{region "05 - Child 1 completes despite the held helper error"}
FSteps[5].Children[1].State := E_State.Completed;
FSteps[5].Children[1].Ready := FALSE;
FSteps[5].Children[1].Complete := TRUE;
FSteps[5].Children[1].Result := E_Result.Passed;
FSteps[5].Children[2].State := E_State.Idle;
FSteps[5].Children[2].Ready := FALSE;
FSteps[5].ExpectedSlot := 1;
FSteps[5].ExpectedReservations[1] := 1;
FSteps[5].MaxActiveChildCount := 1;
FSteps[5].ExpectedResult := E_Result.Error;
FSteps[5].ExpectedDiagnosticCount := 1;
{endregion}

{region "06 - Release the completed child only"}
FSteps[6].Children[1].State := E_State.Completed;
FSteps[6].Children[1].Ready := FALSE;
FSteps[6].Children[1].Complete := TRUE;
FSteps[6].Children[1].Result := E_Result.Passed;
FSteps[6].Children[2].State := E_State.Idle;
FSteps[6].Children[2].Ready := FALSE;
FSteps[6].ExpectedSlot := 1;
FSteps[6].ExpectedReleasedEntries[1] := 1;
FSteps[6].MaxActiveChildCount := 0;
FSteps[6].ExpectedResult := E_Result.Error;
FSteps[6].ExpectedDiagnosticCount := 1;
{endregion}

{region "07 - Readiness recovery does not clear the held error"}
FSteps[7].Children[1].State := E_State.Completed;
FSteps[7].Children[1].Ready := FALSE;
FSteps[7].Children[1].Complete := TRUE;
FSteps[7].Children[1].Result := E_Result.Passed;
FSteps[7].ExpectedSlot := 1;
FSteps[7].MaxActiveChildCount := 0;
FSteps[7].ExpectedResult := E_Result.Error;
FSteps[7].ExpectedDiagnosticCount := 1;
{endregion}

{region "08 - Recovered readiness cannot restart execution"}
FSteps[8].Children[1].State := E_State.Completed;
FSteps[8].Children[1].Ready := FALSE;
FSteps[8].Children[1].Complete := TRUE;
FSteps[8].Children[1].Result := E_Result.Passed;
FSteps[8].ExpectedSlot := 1;
FSteps[8].MaxActiveChildCount := 0;
FSteps[8].ExpectedResult := E_Result.Error;
FSteps[8].ExpectedDiagnosticCount := 1;
{endregion}
END_METHOD

END_FUNCTION_BLOCK

// ---- SelfTests/TestCases/TestSuite_ParallelOrchestration/Test_ParallelFailedResultContinues.TcPOU
{region 'Documentation'}
(*!
<summary>Keeps parallel siblings progressing after a child completes with Failed instead of treating it as a helper Error.</summary>
<description>
Child 1 finishes with Failed while child 2 starts. Child 3 must still start while child 2
runs. The helper reports neutral Result and completes only after all children;
child-result aggregation belongs to the owner.
</description>
*)
{endregion}
FUNCTION_BLOCK Test_ParallelFailedResultContinues EXTENDS OrchestrationTestBase

SUPER^();

{region 'Documentation'}
(*!
<summary>Defines reachable child responses and independent per-cycle expectations.</summary>
*)
{endregion}
METHOD PROTECTED ConfigureScenario
FChildSlots[1] := 1;
FChildSlots[2] := 1;
FChildSlots[3] := 1;
FStepCount := 7;

{region "01 - Observe initial readiness"}
FSteps[1].Task := E_OrchestratorTask.Idle;
FSteps[1].ExpectedReady := TRUE;
{endregion}

{region "02 - Start child 1"}
FSteps[2].Children[1].State := E_State.Running;
FSteps[2].Children[1].Ready := FALSE;
FSteps[2].ExpectedStartChild := 1;
FSteps[2].ExpectedSlot := 1;
FSteps[2].ExpectedReservations[1] := 1;
FSteps[2].MaxActiveChildCount := 1;
{endregion}

{region "03 - Start child 2 while child 1 finishes with Failed"}
FSteps[3].Children[1].State := E_State.Completed;
FSteps[3].Children[1].Ready := FALSE;
FSteps[3].Children[1].Complete := TRUE;
FSteps[3].Children[1].Result := E_Result.Failed;
FSteps[3].Children[2].State := E_State.Running;
FSteps[3].Children[2].Ready := FALSE;
FSteps[3].ExpectedStartChild := 2;
FSteps[3].ExpectedSlot := 1;
FSteps[3].ExpectedReservations[1] := 1;
FSteps[3].ExpectedReservations[2] := 1;
FSteps[3].MaxActiveChildCount := 2;
{endregion}

{region "04 - Release Failed child 1 and start child 3"}
FSteps[4].Children[1].State := E_State.Completed;
FSteps[4].Children[1].Ready := FALSE;
FSteps[4].Children[1].Complete := TRUE;
FSteps[4].Children[1].Result := E_Result.Failed;
FSteps[4].Children[2].State := E_State.Running;
FSteps[4].Children[2].Ready := FALSE;
FSteps[4].Children[3].State := E_State.Running;
FSteps[4].Children[3].Ready := FALSE;
FSteps[4].ExpectedStartChild := 3;
FSteps[4].ExpectedSlot := 1;
FSteps[4].ExpectedReservations[2] := 1;
FSteps[4].ExpectedReservations[3] := 1;
FSteps[4].ExpectedReleasedEntries[1] := 1;
FSteps[4].MaxActiveChildCount := 2;
{endregion}

{region "05 - Remaining children complete without helper Error"}
FSteps[5].Children[1].State := E_State.Completed;
FSteps[5].Children[1].Ready := FALSE;
FSteps[5].Children[1].Complete := TRUE;
FSteps[5].Children[1].Result := E_Result.Failed;
FSteps[5].Children[2].State := E_State.Completed;
FSteps[5].Children[2].Ready := FALSE;
FSteps[5].Children[2].Complete := TRUE;
FSteps[5].Children[2].Result := E_Result.Passed;
FSteps[5].Children[3].State := E_State.Completed;
FSteps[5].Children[3].Ready := FALSE;
FSteps[5].Children[3].Complete := TRUE;
FSteps[5].Children[3].Result := E_Result.Passed;
FSteps[5].ExpectedSlot := 1;
FSteps[5].ExpectedReservations[2] := 1;
FSteps[5].ExpectedReservations[3] := 1;
FSteps[5].MaxActiveChildCount := 2;
{endregion}

{region "06 - Release both siblings and finish the whole group"}
FSteps[6].Children[1].State := E_State.Completed;
FSteps[6].Children[1].Ready := FALSE;
FSteps[6].Children[1].Complete := TRUE;
FSteps[6].Children[1].Result := E_Result.Failed;
FSteps[6].Children[2].State := E_State.Completed;
FSteps[6].Children[2].Ready := FALSE;
FSteps[6].Children[2].Complete := TRUE;
FSteps[6].Children[2].Result := E_Result.Passed;
FSteps[6].Children[3].State := E_State.Completed;
FSteps[6].Children[3].Ready := FALSE;
FSteps[6].Children[3].Complete := TRUE;
FSteps[6].Children[3].Result := E_Result.Passed;
FSteps[6].ExpectedFinished := TRUE;
FSteps[6].ExpectedReleasedEntries[2] := 1;
FSteps[6].ExpectedReleasedEntries[3] := 1;
FSteps[6].MaxActiveChildCount := 0;
{endregion}

{region "07 - Keep completion stable with neutral helper Result"}
FSteps[7].Children[1].State := E_State.Completed;
FSteps[7].Children[1].Ready := FALSE;
FSteps[7].Children[1].Complete := TRUE;
FSteps[7].Children[1].Result := E_Result.Failed;
FSteps[7].Children[2].State := E_State.Completed;
FSteps[7].Children[2].Ready := FALSE;
FSteps[7].Children[2].Complete := TRUE;
FSteps[7].Children[2].Result := E_Result.Passed;
FSteps[7].Children[3].State := E_State.Completed;
FSteps[7].Children[3].Ready := FALSE;
FSteps[7].Children[3].Complete := TRUE;
FSteps[7].Children[3].Result := E_Result.Passed;
FSteps[7].ExpectedFinished := TRUE;
FSteps[7].MaxActiveChildCount := 0;
{endregion}
END_METHOD

END_FUNCTION_BLOCK

// ---- SelfTests/TestCases/TestSuite_ParallelOrchestration/Test_ParallelChildError.TcPOU
{region 'Documentation'}
(*!
<summary>Stops new parallel Starts on child Error and observes owner-selected Abort of the remaining active sibling.</summary>
<description>
Child 1 enters its error-abort path while child 2 starts. The helper must retain Error and
not start child 3. The owner then supplies Abort explicitly; already-aborting child 1 and
never-started child 3 receive no redundant Abort.
</description>
*)
{endregion}
FUNCTION_BLOCK Test_ParallelChildError EXTENDS OrchestrationTestBase

SUPER^();

{region 'Documentation'}
(*!
<summary>Defines reachable child responses and independent per-cycle expectations.</summary>
*)
{endregion}
METHOD PROTECTED ConfigureScenario
FChildSlots[1] := 1;
FChildSlots[2] := 1;
FChildSlots[3] := 1;
FStepCount := 8;

{region "01 - Observe initial readiness"}
FSteps[1].Task := E_OrchestratorTask.Idle;
FSteps[1].ExpectedReady := TRUE;
{endregion}

{region "02 - Start child 1 normally"}
FSteps[2].Children[1].State := E_State.Running;
FSteps[2].Children[1].Ready := FALSE;
FSteps[2].ExpectedStartChild := 1;
FSteps[2].ExpectedSlot := 1;
FSteps[2].ExpectedReservations[1] := 1;
FSteps[2].MaxActiveChildCount := 1;
{endregion}

{region "03 - Start child 2 while child 1 enters its error path"}
FSteps[3].Children[1].State := E_State.AbortingFromError;
FSteps[3].Children[1].Ready := FALSE;
FSteps[3].Children[1].Result := E_Result.Error;
FSteps[3].Children[2].State := E_State.Running;
FSteps[3].Children[2].Ready := FALSE;
FSteps[3].ExpectedStartChild := 2;
FSteps[3].ExpectedSlot := 1;
FSteps[3].ExpectedReservations[1] := 1;
FSteps[3].ExpectedReservations[2] := 1;
FSteps[3].MaxActiveChildCount := 2;
{endregion}

{region "04 - Observe child Error and suppress child 3 Start"}
FSteps[4].Children[1].State := E_State.AbortingFromError;
FSteps[4].Children[1].Ready := FALSE;
FSteps[4].Children[1].Result := E_Result.Error;
FSteps[4].Children[2].State := E_State.Running;
FSteps[4].Children[2].Ready := FALSE;
FSteps[4].ExpectedSlot := 1;
FSteps[4].ExpectedReservations[1] := 1;
FSteps[4].ExpectedReservations[2] := 1;
FSteps[4].MaxActiveChildCount := 2;
FSteps[4].ExpectedResult := E_Result.Error;
FSteps[4].ExpectedDiagnosticCount := 1;
{endregion}

{region "05 - Owner selects Abort for remaining active work"}
FSteps[5].Task := E_OrchestratorTask.Abort;
FSteps[5].Children[1].State := E_State.AbortingFromError;
FSteps[5].Children[1].Ready := FALSE;
FSteps[5].Children[1].Result := E_Result.Error;
FSteps[5].Children[2].State := E_State.Aborting;
FSteps[5].Children[2].Ready := FALSE;
FSteps[5].Children[2].Result := E_Result.Abort;
FSteps[5].ExpectedReservations[1] := 1;
FSteps[5].ExpectedReservations[2] := 1;
FSteps[5].ExpectedAbortRequests[2] := 1;
FSteps[5].ExpectedResult := E_Result.Error;
FSteps[5].ExpectedDiagnosticCount := 1;
{endregion}

{region "06 - Both active children reach terminal states"}
FSteps[6].Task := E_OrchestratorTask.Abort;
FSteps[6].Children[1].State := E_State.Completed;
FSteps[6].Children[1].Ready := FALSE;
FSteps[6].Children[1].Complete := TRUE;
FSteps[6].Children[1].Result := E_Result.Error;
FSteps[6].Children[2].State := E_State.Completed;
FSteps[6].Children[2].Ready := FALSE;
FSteps[6].Children[2].Complete := TRUE;
FSteps[6].Children[2].Result := E_Result.Abort;
FSteps[6].ExpectedReservations[1] := 1;
FSteps[6].ExpectedReservations[2] := 1;
FSteps[6].ExpectedResult := E_Result.Error;
FSteps[6].ExpectedDiagnosticCount := 1;
{endregion}

{region "07 - Release terminal reservations and finish Abort"}
FSteps[7].Task := E_OrchestratorTask.Abort;
FSteps[7].Children[1].State := E_State.Completed;
FSteps[7].Children[1].Ready := FALSE;
FSteps[7].Children[1].Complete := TRUE;
FSteps[7].Children[1].Result := E_Result.Error;
FSteps[7].Children[2].State := E_State.Completed;
FSteps[7].Children[2].Ready := FALSE;
FSteps[7].Children[2].Complete := TRUE;
FSteps[7].Children[2].Result := E_Result.Abort;
FSteps[7].ExpectedAbortFinished := TRUE;
FSteps[7].ExpectedReleasedEntries[1] := 1;
FSteps[7].ExpectedReleasedEntries[2] := 1;
FSteps[7].ExpectedResult := E_Result.Error;
FSteps[7].ExpectedDiagnosticCount := 1;
{endregion}

{region "08 - Repeated Abort neither redispatches nor republishes"}
FSteps[8].Task := E_OrchestratorTask.Abort;
FSteps[8].Children[1].State := E_State.Completed;
FSteps[8].Children[1].Ready := FALSE;
FSteps[8].Children[1].Complete := TRUE;
FSteps[8].Children[1].Result := E_Result.Error;
FSteps[8].Children[2].State := E_State.Completed;
FSteps[8].Children[2].Ready := FALSE;
FSteps[8].Children[2].Complete := TRUE;
FSteps[8].Children[2].Result := E_Result.Abort;
FSteps[8].ExpectedAbortFinished := TRUE;
FSteps[8].ExpectedResult := E_Result.Error;
FSteps[8].ExpectedDiagnosticCount := 1;
{endregion}
END_METHOD

END_FUNCTION_BLOCK

// ---- SelfTests/TestCases/TestSuite_ParallelOrchestration/Test_ParallelAbortMixedProgress.TcPOU
{region 'Documentation'}
(*!
<summary>Aborts only active parallel work while leaving completed and never-started ready children untouched.</summary>
<description>
Child 2 completes on its Start call while child 1 runs. The owner selects Abort before
child 3 starts. Start confirmation, terminal release and active-child Abort happen in the
same helper call; completion waits for child 1.
</description>
*)
{endregion}
FUNCTION_BLOCK Test_ParallelAbortMixedProgress EXTENDS OrchestrationTestBase

SUPER^();

{region 'Documentation'}
(*!
<summary>Defines reachable child responses and independent per-cycle expectations.</summary>
*)
{endregion}
METHOD PROTECTED ConfigureScenario
FChildSlots[1] := 1;
FChildSlots[2] := 1;
FChildSlots[3] := 1;
FStepCount := 7;

{region "01 - Observe initial readiness"}
FSteps[1].Task := E_OrchestratorTask.Idle;
FSteps[1].ExpectedReady := TRUE;
{endregion}

{region "02 - Start child 1"}
FSteps[2].Children[1].State := E_State.Running;
FSteps[2].Children[1].Ready := FALSE;
FSteps[2].ExpectedStartChild := 1;
FSteps[2].ExpectedSlot := 1;
FSteps[2].ExpectedReservations[1] := 1;
FSteps[2].MaxActiveChildCount := 1;
{endregion}

{region "03 - Start immediately completing child 2"}
FSteps[3].Children[1].State := E_State.Running;
FSteps[3].Children[1].Ready := FALSE;
FSteps[3].Children[2].State := E_State.Completed;
FSteps[3].Children[2].Ready := FALSE;
FSteps[3].Children[2].Complete := TRUE;
FSteps[3].Children[2].Result := E_Result.Passed;
FSteps[3].ExpectedStartChild := 2;
FSteps[3].ExpectedSlot := 1;
FSteps[3].ExpectedReservations[1] := 1;
FSteps[3].ExpectedReservations[2] := 1;
FSteps[3].MaxActiveChildCount := 2;
{endregion}

{region "04 - Owner selects Abort while child 3 remains unstarted"}
FSteps[4].Task := E_OrchestratorTask.Abort;
FSteps[4].Children[1].State := E_State.Aborting;
FSteps[4].Children[1].Ready := FALSE;
FSteps[4].Children[1].Result := E_Result.Abort;
FSteps[4].Children[2].State := E_State.Completed;
FSteps[4].Children[2].Ready := FALSE;
FSteps[4].Children[2].Complete := TRUE;
FSteps[4].Children[2].Result := E_Result.Passed;
FSteps[4].ExpectedReservations[1] := 1;
FSteps[4].ExpectedReleasedEntries[2] := 1;
FSteps[4].ExpectedAbortRequests[1] := 1;
{endregion}

{region "05 - Wait for the active child's controlled completion"}
FSteps[5].Task := E_OrchestratorTask.Abort;
FSteps[5].Children[1].State := E_State.Completed;
FSteps[5].Children[1].Ready := FALSE;
FSteps[5].Children[1].Complete := TRUE;
FSteps[5].Children[1].Result := E_Result.Abort;
FSteps[5].Children[2].State := E_State.Completed;
FSteps[5].Children[2].Ready := FALSE;
FSteps[5].Children[2].Complete := TRUE;
FSteps[5].Children[2].Result := E_Result.Passed;
FSteps[5].ExpectedReservations[1] := 1;
{endregion}

{region "06 - Release child 1 and finish Abort"}
FSteps[6].Task := E_OrchestratorTask.Abort;
FSteps[6].Children[1].State := E_State.Completed;
FSteps[6].Children[1].Ready := FALSE;
FSteps[6].Children[1].Complete := TRUE;
FSteps[6].Children[1].Result := E_Result.Abort;
FSteps[6].Children[2].State := E_State.Completed;
FSteps[6].Children[2].Ready := FALSE;
FSteps[6].Children[2].Complete := TRUE;
FSteps[6].Children[2].Result := E_Result.Passed;
FSteps[6].ExpectedAbortFinished := TRUE;
FSteps[6].ExpectedReleasedEntries[1] := 1;
{endregion}

{region "07 - No repeated Abort or new Start after completion"}
FSteps[7].Task := E_OrchestratorTask.Abort;
FSteps[7].Children[1].State := E_State.Completed;
FSteps[7].Children[1].Ready := FALSE;
FSteps[7].Children[1].Complete := TRUE;
FSteps[7].Children[1].Result := E_Result.Abort;
FSteps[7].Children[2].State := E_State.Completed;
FSteps[7].Children[2].Ready := FALSE;
FSteps[7].Children[2].Complete := TRUE;
FSteps[7].Children[2].Result := E_Result.Passed;
FSteps[7].ExpectedAbortFinished := TRUE;
{endregion}
END_METHOD

END_FUNCTION_BLOCK

// ---- SelfTests/TestCases/TestSuite_ParallelOrchestration/Test_ParallelResetOverlappingExecution.TcPOU
{region 'Documentation'}
(*!
<summary>Resets overlapping parallel children and an already completed child without issuing further Starts.</summary>
<description>
Two children are running when the third completes immediately. Owner-selected Reset
replaces each execution reservation through the child's Reset reservation method.
Independent reset completion retains unfinished reservations and returns to ready Idle
only after all children finish.
</description>
*)
{endregion}
FUNCTION_BLOCK Test_ParallelResetOverlappingExecution EXTENDS OrchestrationTestBase

SUPER^();

{region 'Documentation'}
(*!
<summary>Defines reachable child responses and independent per-cycle expectations.</summary>
*)
{endregion}
METHOD PROTECTED ConfigureScenario
FChildSlots[1] := 1;
FChildSlots[2] := 1;
FChildSlots[3] := 1;
FStepCount := 12;

{region "01 - Observe initial readiness"}
FSteps[1].Task := E_OrchestratorTask.Idle;
FSteps[1].ExpectedReady := TRUE;
{endregion}

{region "02 - Start child 1"}
FSteps[2].Children[1].State := E_State.Running;
FSteps[2].Children[1].Ready := FALSE;
FSteps[2].ExpectedStartChild := 1;
FSteps[2].ExpectedSlot := 1;
FSteps[2].ExpectedReservations[1] := 1;
FSteps[2].MaxActiveChildCount := 1;
{endregion}

{region "03 - Start child 2 concurrently"}
FSteps[3].Children[1].State := E_State.Running;
FSteps[3].Children[1].Ready := FALSE;
FSteps[3].Children[2].State := E_State.Running;
FSteps[3].Children[2].Ready := FALSE;
FSteps[3].ExpectedStartChild := 2;
FSteps[3].ExpectedSlot := 1;
FSteps[3].ExpectedReservations[1] := 1;
FSteps[3].ExpectedReservations[2] := 1;
FSteps[3].MaxActiveChildCount := 2;
{endregion}

{region "04 - Start child 3 which completes immediately"}
FSteps[4].Children[1].State := E_State.Running;
FSteps[4].Children[1].Ready := FALSE;
FSteps[4].Children[2].State := E_State.Running;
FSteps[4].Children[2].Ready := FALSE;
FSteps[4].Children[3].State := E_State.Completed;
FSteps[4].Children[3].Ready := FALSE;
FSteps[4].Children[3].Complete := TRUE;
FSteps[4].Children[3].Result := E_Result.Passed;
FSteps[4].ExpectedStartChild := 3;
FSteps[4].ExpectedSlot := 1;
FSteps[4].ExpectedReservations[1] := 1;
FSteps[4].ExpectedReservations[2] := 1;
FSteps[4].ExpectedReservations[3] := 1;
FSteps[4].MaxActiveChildCount := 3;
{endregion}

{region "05 - Owner selects Reset and resets active child 1"}
FSteps[5].Task := E_OrchestratorTask.Reset;
FSteps[5].Children[1].State := E_State.Reset;
FSteps[5].Children[1].Ready := FALSE;
FSteps[5].Children[2].State := E_State.Running;
FSteps[5].Children[2].Ready := FALSE;
FSteps[5].Children[3].State := E_State.Completed;
FSteps[5].Children[3].Ready := FALSE;
FSteps[5].Children[3].Complete := TRUE;
FSteps[5].Children[3].Result := E_Result.Passed;
FSteps[5].ExpectedResetChild := 1;
FSteps[5].ExpectedReservations[1] := 1;
FSteps[5].ExpectedReservations[2] := 1;
FSteps[5].ExpectedReservations[3] := 1;
{endregion}

{region "06 - Reset child 2 while child 1 is still resetting"}
FSteps[6].Task := E_OrchestratorTask.Reset;
FSteps[6].Children[1].State := E_State.Reset;
FSteps[6].Children[1].Ready := FALSE;
FSteps[6].Children[2].State := E_State.Reset;
FSteps[6].Children[2].Ready := FALSE;
FSteps[6].Children[3].State := E_State.Completed;
FSteps[6].Children[3].Ready := FALSE;
FSteps[6].Children[3].Complete := TRUE;
FSteps[6].Children[3].Result := E_Result.Passed;
FSteps[6].ExpectedResetChild := 2;
FSteps[6].ExpectedReservations[1] := 1;
FSteps[6].ExpectedReservations[2] := 1;
FSteps[6].ExpectedReservations[3] := 1;
{endregion}

{region "07 - Reset completed child 3 while child 1 reaches Idle"}
FSteps[7].Task := E_OrchestratorTask.Reset;
FSteps[7].Children[2].State := E_State.Reset;
FSteps[7].Children[2].Ready := FALSE;
FSteps[7].Children[3].State := E_State.Reset;
FSteps[7].Children[3].Ready := FALSE;
FSteps[7].ExpectedResetChild := 3;
FSteps[7].ExpectedReservations[1] := 1;
FSteps[7].ExpectedReservations[2] := 1;
FSteps[7].ExpectedReservations[3] := 1;
{endregion}

{region "08 - Release child 1 while child 2 reaches Idle"}
FSteps[8].Task := E_OrchestratorTask.Reset;
FSteps[8].Children[3].State := E_State.Reset;
FSteps[8].Children[3].Ready := FALSE;
FSteps[8].ExpectedReservations[2] := 1;
FSteps[8].ExpectedReservations[3] := 1;
FSteps[8].ExpectedReleasedEntries[1] := 1;
{endregion}

{region "09 - Release child 2 while child 3 reaches Idle"}
FSteps[9].Task := E_OrchestratorTask.Reset;
FSteps[9].ExpectedReservations[3] := 1;
FSteps[9].ExpectedReleasedEntries[2] := 1;
{endregion}

{region "10 - Release final reservation and report Reset finished"}
FSteps[10].Task := E_OrchestratorTask.Reset;
FSteps[10].ExpectedResetFinished := TRUE;
FSteps[10].ExpectedReleasedEntries[3] := 1;
{endregion}

{region "11 - Repeated Reset retains completion without redispatch"}
FSteps[11].Task := E_OrchestratorTask.Reset;
FSteps[11].ExpectedResetFinished := TRUE;
{endregion}

{region "12 - Owner selects Idle and observes restored readiness"}
FSteps[12].Task := E_OrchestratorTask.Idle;
FSteps[12].ExpectedReady := TRUE;
{endregion}
END_METHOD

END_FUNCTION_BLOCK

// ---- SelfTests/TestSuites/TestSuite_ParallelSlotsOrchestration.TcPOU
{region 'Documentation'}
(*!
<summary>Runs focused ParallelSlots Orchestrator scenarios serially with isolated child observations and diagnostics.</summary>
*)
{endregion}
FUNCTION_BLOCK TestSuite_ParallelSlotsOrchestration EXTENDS TestSuiteBase
VAR
    FWaitForGroupCompletion : Test_SlotsWaitForGroupCompletion;
    FFinalGroupCompletion : Test_SlotsFinalGroupCompletion;
    FFirstFittingAdmission : Test_SlotsFirstFittingAdmission;
    FMissingStartReaction : Test_SlotsMissingStartReaction;
    FNextSlotReadinessLost : Test_SlotsNextSlotReadinessLost;
    FAbortAtBoundary : Test_SlotsAbortAtBoundary;
    FTestCases : ARRAY[1..TestCaseCapacity] OF I_TestCase;
END_VAR
VAR CONSTANT
    TestCaseCapacity : UINT := 6;
END_VAR

SUPER^();

{region 'Documentation'}
(*!
<summary>Initializes and registers the owned orchestration scenarios in deterministic order.</summary>
*)
{endregion}
METHOD PROTECTED Configure
VAR_IN_OUT
    // SA0167: Borrowed builder; VAR_IN_OUT creates no temporary instance.
    {attribute 'analysis' := '-167'}
    Builder : TestSuiteConfigurationBuilder; //! Borrowed owner configuration builder used only during this Configure call; register this owner's concrete children.
END_VAR
VAR
    TestConfig : ST_TestCaseConfig;
END_VAR
Builder.Initialize(Mode := E_OrchestrationMode.Serial,
    TestCases := FTestCases);

FWaitForGroupCompletion.Initialize(Parent := THIS^,
    TestName := 'WaitForGroupCompletion',
    Config := TestConfig);
Builder.Register(TestCase := FWaitForGroupCompletion);

FFinalGroupCompletion.Initialize(Parent := THIS^,
    TestName := 'FinalGroupCompletion',
    Config := TestConfig);
Builder.Register(TestCase := FFinalGroupCompletion);

FFirstFittingAdmission.Initialize(Parent := THIS^,
    TestName := 'FirstFittingAdmission',
    Config := TestConfig);
Builder.Register(TestCase := FFirstFittingAdmission);

FMissingStartReaction.Initialize(Parent := THIS^,
    TestName := 'MissingStartReaction',
    Config := TestConfig);
Builder.Register(TestCase := FMissingStartReaction);

FNextSlotReadinessLost.Initialize(Parent := THIS^,
    TestName := 'NextSlotReadinessLost',
    Config := TestConfig);
Builder.Register(TestCase := FNextSlotReadinessLost);

FAbortAtBoundary.Initialize(Parent := THIS^,
    TestName := 'AbortAtBoundary',
    Config := TestConfig);
Builder.Register(TestCase := FAbortAtBoundary);
END_METHOD

{region 'Documentation'}
(*!
<summary>Returns the registered Test Case from the same array used during configuration.</summary>
*)
{endregion}
METHOD PUBLIC GetTestCase : I_TestCase //! Typed child interface at the original array index; zero when no entry is available.
VAR_INPUT
    Index : DINT; //! Original occupied child-array index, rather than an ordinal position.
END_VAR
GetTestCase := 0;
IF (ChildCount = 0) OR (Index < ChildArrayLowerBound)
    OR (DINT_TO_LINT(Index) >= DINT_TO_LINT(ChildArrayLowerBound) + UINT_TO_LINT(ChildCount)) THEN
    RETURN;
END_IF;

GetTestCase := FTestCases[Index];
END_METHOD

{region 'Documentation'}
(*!
<summary>Calls each owned Test Case once per initialized Suite cycle, including completion.</summary>
*)
{endregion}
METHOD PROTECTED ProcessTestCases
FWaitForGroupCompletion();
FFinalGroupCompletion();
FFirstFittingAdmission();
FMissingStartReaction();
FNextSlotReadinessLost();
FAbortAtBoundary();
END_METHOD

END_FUNCTION_BLOCK

// ---- SelfTests/TestCases/TestSuite_ParallelSlotsOrchestration/Test_SlotsWaitForGroupCompletion.TcPOU
{region 'Documentation'}
(*!
<summary>Keeps the next slot blocked until both unequal-duration children in the current slot complete.</summary>
<description>
Children 1 and 2 share slot 1. Child 2 finishes first while child 1 remains active.
Child 3 stays idle in slot 2 until both earlier children complete and their reservations
are released. Each row observes the helper before applying the next child responses.
</description>
*)
{endregion}
FUNCTION_BLOCK Test_SlotsWaitForGroupCompletion EXTENDS OrchestrationTestBase

SUPER^();

{region 'Documentation'}
(*!
<summary>Defines slot-group stimuli and per-cycle dispatch, completion and reservation expectations.</summary>
*)
{endregion}
METHOD PROTECTED ConfigureScenario
FChildSlots[1] := 1;
FChildSlots[2] := 1;
FChildSlots[3] := 2;
FStepCount := 11;

{region "01 - Observe initial readiness"}
FSteps[1].Task := E_OrchestratorTask.Idle;
FSteps[1].ExpectedReady := TRUE;
FSteps[1].MaxActiveChildCount := 0;
{endregion}

{region "02 - Start long-running child 1 in slot 1"}
FSteps[2].Children[1].State := E_State.Running;
FSteps[2].Children[1].Ready := FALSE;
FSteps[2].ExpectedStartChild := 1;
FSteps[2].ExpectedSlot := 1;
FSteps[2].ExpectedReservations[1] := 1;
FSteps[2].MaxActiveChildCount := 1;
{endregion}

{region "03 - Start child 2 alongside child 1"}
FSteps[3].Children[1].State := E_State.Running;
FSteps[3].Children[1].Ready := FALSE;
FSteps[3].Children[2].State := E_State.Running;
FSteps[3].Children[2].Ready := FALSE;
FSteps[3].ExpectedStartChild := 2;
FSteps[3].ExpectedSlot := 1;
FSteps[3].ExpectedReservations[1] := 1;
FSteps[3].ExpectedReservations[2] := 1;
FSteps[3].MaxActiveChildCount := 2;
{endregion}

{region "04 - Child 2 completes while child 1 remains active"}
FSteps[4].Children[1].State := E_State.Running;
FSteps[4].Children[1].Ready := FALSE;
FSteps[4].Children[2].State := E_State.Completed;
FSteps[4].Children[2].Ready := FALSE;
FSteps[4].Children[2].Complete := TRUE;
FSteps[4].Children[2].Result := E_Result.Passed;
FSteps[4].ExpectedSlot := 1;
FSteps[4].ExpectedReservations[1] := 1;
FSteps[4].ExpectedReservations[2] := 1;
FSteps[4].MaxActiveChildCount := 2;
{endregion}

{region "05 - Release child 2 without starting the next slot"}
FSteps[5].Children[1].State := E_State.Running;
FSteps[5].Children[1].Ready := FALSE;
FSteps[5].Children[2].State := E_State.Completed;
FSteps[5].Children[2].Ready := FALSE;
FSteps[5].Children[2].Complete := TRUE;
FSteps[5].Children[2].Result := E_Result.Passed;
FSteps[5].ExpectedSlot := 1;
FSteps[5].ExpectedReservations[1] := 1;
FSteps[5].ExpectedReleasedEntries[2] := 1;
FSteps[5].MaxActiveChildCount := 1;
{endregion}

{region "06 - Child 1 completes while child 3 still receives no Start"}
FSteps[6].Children[1].State := E_State.Completed;
FSteps[6].Children[1].Ready := FALSE;
FSteps[6].Children[1].Complete := TRUE;
FSteps[6].Children[1].Result := E_Result.Passed;
FSteps[6].Children[2].State := E_State.Completed;
FSteps[6].Children[2].Ready := FALSE;
FSteps[6].Children[2].Complete := TRUE;
FSteps[6].Children[2].Result := E_Result.Passed;
FSteps[6].ExpectedSlot := 1;
FSteps[6].ExpectedReservations[1] := 1;
FSteps[6].MaxActiveChildCount := 1;
{endregion}

{region "07 - Reconcile slot 1 and select slot 2 without dispatch"}
FSteps[7].Children[1].State := E_State.Completed;
FSteps[7].Children[1].Ready := FALSE;
FSteps[7].Children[1].Complete := TRUE;
FSteps[7].Children[1].Result := E_Result.Passed;
FSteps[7].Children[2].State := E_State.Completed;
FSteps[7].Children[2].Ready := FALSE;
FSteps[7].Children[2].Complete := TRUE;
FSteps[7].Children[2].Result := E_Result.Passed;
FSteps[7].ExpectedSlot := 2;
FSteps[7].ExpectedReleasedEntries[1] := 1;
FSteps[7].MaxActiveChildCount := 0;
{endregion}

{region "08 - Start child 3 only after the first group has finished"}
FSteps[8].Children[1].State := E_State.Completed;
FSteps[8].Children[1].Ready := FALSE;
FSteps[8].Children[1].Complete := TRUE;
FSteps[8].Children[1].Result := E_Result.Passed;
FSteps[8].Children[2].State := E_State.Completed;
FSteps[8].Children[2].Ready := FALSE;
FSteps[8].Children[2].Complete := TRUE;
FSteps[8].Children[2].Result := E_Result.Passed;
FSteps[8].Children[3].State := E_State.Running;
FSteps[8].Children[3].Ready := FALSE;
FSteps[8].ExpectedStartChild := 3;
FSteps[8].ExpectedSlot := 2;
FSteps[8].ExpectedReservations[3] := 1;
FSteps[8].MaxActiveChildCount := 1;
{endregion}

{region "09 - Last child completes without redispatching earlier children"}
FSteps[9].Children[1].State := E_State.Completed;
FSteps[9].Children[1].Ready := FALSE;
FSteps[9].Children[1].Complete := TRUE;
FSteps[9].Children[1].Result := E_Result.Passed;
FSteps[9].Children[2].State := E_State.Completed;
FSteps[9].Children[2].Ready := FALSE;
FSteps[9].Children[2].Complete := TRUE;
FSteps[9].Children[2].Result := E_Result.Passed;
FSteps[9].Children[3].State := E_State.Completed;
FSteps[9].Children[3].Ready := FALSE;
FSteps[9].Children[3].Complete := TRUE;
FSteps[9].Children[3].Result := E_Result.Passed;
FSteps[9].ExpectedSlot := 2;
FSteps[9].ExpectedReservations[3] := 1;
FSteps[9].MaxActiveChildCount := 1;
{endregion}

{region "10 - Release the last reservation and finish all slots"}
FSteps[10].Children[1].State := E_State.Completed;
FSteps[10].Children[1].Ready := FALSE;
FSteps[10].Children[1].Complete := TRUE;
FSteps[10].Children[1].Result := E_Result.Passed;
FSteps[10].Children[2].State := E_State.Completed;
FSteps[10].Children[2].Ready := FALSE;
FSteps[10].Children[2].Complete := TRUE;
FSteps[10].Children[2].Result := E_Result.Passed;
FSteps[10].Children[3].State := E_State.Completed;
FSteps[10].Children[3].Ready := FALSE;
FSteps[10].Children[3].Complete := TRUE;
FSteps[10].Children[3].Result := E_Result.Passed;
FSteps[10].ExpectedFinished := TRUE;
FSteps[10].ExpectedReleasedEntries[3] := 1;
FSteps[10].MaxActiveChildCount := 0;
{endregion}

{region "11 - Keep final completion stable without further Starts"}
FSteps[11].Children[1].State := E_State.Completed;
FSteps[11].Children[1].Ready := FALSE;
FSteps[11].Children[1].Complete := TRUE;
FSteps[11].Children[1].Result := E_Result.Passed;
FSteps[11].Children[2].State := E_State.Completed;
FSteps[11].Children[2].Ready := FALSE;
FSteps[11].Children[2].Complete := TRUE;
FSteps[11].Children[2].Result := E_Result.Passed;
FSteps[11].Children[3].State := E_State.Completed;
FSteps[11].Children[3].Ready := FALSE;
FSteps[11].Children[3].Complete := TRUE;
FSteps[11].Children[3].Result := E_Result.Passed;
FSteps[11].ExpectedFinished := TRUE;
FSteps[11].MaxActiveChildCount := 0;
{endregion}
END_METHOD

END_FUNCTION_BLOCK

// ---- SelfTests/TestCases/TestSuite_ParallelSlotsOrchestration/Test_SlotsFinalGroupCompletion.TcPOU
{region 'Documentation'}
(*!
<summary>Runs both final-slot children in parallel and ignores unused collection capacity when determining completion.</summary>
<description>
Child 1 completes immediately in slot 1. Children 2 and 3 then overlap in the final
slot and finish in reverse order. The collection has six array positions but only three
registered children; final-slot detection must use the occupied range.
</description>
*)
{endregion}
FUNCTION_BLOCK Test_SlotsFinalGroupCompletion EXTENDS OrchestrationTestBase

SUPER^();

{region 'Documentation'}
(*!
<summary>Defines slot-group stimuli and per-cycle dispatch, completion and reservation expectations.</summary>
*)
{endregion}
METHOD PROTECTED ConfigureScenario
FChildSlots[1] := 1;
FChildSlots[2] := 2;
FChildSlots[3] := 2;
FArrayLayout := E_OrchestrationArrayLayout.SpareCapacity;
FStepCount := 10;

{region "01 - Observe readiness with unused array capacity"}
FSteps[1].Task := E_OrchestratorTask.Idle;
FSteps[1].ExpectedReady := TRUE;
FSteps[1].MaxActiveChildCount := 0;
{endregion}

{region "02 - Start child 1 which completes immediately"}
FSteps[2].Children[1].State := E_State.Completed;
FSteps[2].Children[1].Ready := FALSE;
FSteps[2].Children[1].Complete := TRUE;
FSteps[2].Children[1].Result := E_Result.Passed;
FSteps[2].ExpectedStartChild := 1;
FSteps[2].ExpectedSlot := 1;
FSteps[2].ExpectedReservations[1] := 1;
FSteps[2].MaxActiveChildCount := 1;
{endregion}

{region "03 - Confirm immediate completion and select the final slot"}
FSteps[3].Children[1].State := E_State.Completed;
FSteps[3].Children[1].Ready := FALSE;
FSteps[3].Children[1].Complete := TRUE;
FSteps[3].Children[1].Result := E_Result.Passed;
FSteps[3].ExpectedSlot := 2;
FSteps[3].ExpectedReleasedEntries[1] := 1;
FSteps[3].MaxActiveChildCount := 0;
{endregion}

{region "04 - Start child 2 in the final slot"}
FSteps[4].Children[1].State := E_State.Completed;
FSteps[4].Children[1].Ready := FALSE;
FSteps[4].Children[1].Complete := TRUE;
FSteps[4].Children[1].Result := E_Result.Passed;
FSteps[4].Children[2].State := E_State.Running;
FSteps[4].Children[2].Ready := FALSE;
FSteps[4].ExpectedStartChild := 2;
FSteps[4].ExpectedSlot := 2;
FSteps[4].ExpectedReservations[2] := 1;
FSteps[4].MaxActiveChildCount := 1;
{endregion}

{region "05 - Start child 3 while child 2 remains active"}
FSteps[5].Children[1].State := E_State.Completed;
FSteps[5].Children[1].Ready := FALSE;
FSteps[5].Children[1].Complete := TRUE;
FSteps[5].Children[1].Result := E_Result.Passed;
FSteps[5].Children[2].State := E_State.Running;
FSteps[5].Children[2].Ready := FALSE;
FSteps[5].Children[3].State := E_State.Running;
FSteps[5].Children[3].Ready := FALSE;
FSteps[5].ExpectedStartChild := 3;
FSteps[5].ExpectedSlot := 2;
FSteps[5].ExpectedReservations[2] := 1;
FSteps[5].ExpectedReservations[3] := 1;
FSteps[5].MaxActiveChildCount := 2;
{endregion}

{region "06 - Child 3 completes before child 2"}
FSteps[6].Children[1].State := E_State.Completed;
FSteps[6].Children[1].Ready := FALSE;
FSteps[6].Children[1].Complete := TRUE;
FSteps[6].Children[1].Result := E_Result.Passed;
FSteps[6].Children[2].State := E_State.Running;
FSteps[6].Children[2].Ready := FALSE;
FSteps[6].Children[3].State := E_State.Completed;
FSteps[6].Children[3].Ready := FALSE;
FSteps[6].Children[3].Complete := TRUE;
FSteps[6].Children[3].Result := E_Result.Passed;
FSteps[6].ExpectedSlot := 2;
FSteps[6].ExpectedReservations[2] := 1;
FSteps[6].ExpectedReservations[3] := 1;
FSteps[6].MaxActiveChildCount := 2;
{endregion}

{region "07 - Release child 3 without reporting final completion"}
FSteps[7].Children[1].State := E_State.Completed;
FSteps[7].Children[1].Ready := FALSE;
FSteps[7].Children[1].Complete := TRUE;
FSteps[7].Children[1].Result := E_Result.Passed;
FSteps[7].Children[2].State := E_State.Running;
FSteps[7].Children[2].Ready := FALSE;
FSteps[7].Children[3].State := E_State.Completed;
FSteps[7].Children[3].Ready := FALSE;
FSteps[7].Children[3].Complete := TRUE;
FSteps[7].Children[3].Result := E_Result.Passed;
FSteps[7].ExpectedSlot := 2;
FSteps[7].ExpectedReservations[2] := 1;
FSteps[7].ExpectedReleasedEntries[3] := 1;
FSteps[7].MaxActiveChildCount := 1;
{endregion}

{region "08 - Child 2 completes after its shorter sibling"}
FSteps[8].Children[1].State := E_State.Completed;
FSteps[8].Children[1].Ready := FALSE;
FSteps[8].Children[1].Complete := TRUE;
FSteps[8].Children[1].Result := E_Result.Passed;
FSteps[8].Children[2].State := E_State.Completed;
FSteps[8].Children[2].Ready := FALSE;
FSteps[8].Children[2].Complete := TRUE;
FSteps[8].Children[2].Result := E_Result.Passed;
FSteps[8].Children[3].State := E_State.Completed;
FSteps[8].Children[3].Ready := FALSE;
FSteps[8].Children[3].Complete := TRUE;
FSteps[8].Children[3].Result := E_Result.Passed;
FSteps[8].ExpectedSlot := 2;
FSteps[8].ExpectedReservations[2] := 1;
FSteps[8].MaxActiveChildCount := 1;
{endregion}

{region "09 - Finish at the occupied boundary rather than array capacity"}
FSteps[9].Children[1].State := E_State.Completed;
FSteps[9].Children[1].Ready := FALSE;
FSteps[9].Children[1].Complete := TRUE;
FSteps[9].Children[1].Result := E_Result.Passed;
FSteps[9].Children[2].State := E_State.Completed;
FSteps[9].Children[2].Ready := FALSE;
FSteps[9].Children[2].Complete := TRUE;
FSteps[9].Children[2].Result := E_Result.Passed;
FSteps[9].Children[3].State := E_State.Completed;
FSteps[9].Children[3].Ready := FALSE;
FSteps[9].Children[3].Complete := TRUE;
FSteps[9].Children[3].Result := E_Result.Passed;
FSteps[9].ExpectedFinished := TRUE;
FSteps[9].ExpectedReleasedEntries[2] := 1;
FSteps[9].MaxActiveChildCount := 0;
{endregion}

{region "10 - Keep completion stable without accessing spare entries"}
FSteps[10].Children[1].State := E_State.Completed;
FSteps[10].Children[1].Ready := FALSE;
FSteps[10].Children[1].Complete := TRUE;
FSteps[10].Children[1].Result := E_Result.Passed;
FSteps[10].Children[2].State := E_State.Completed;
FSteps[10].Children[2].Ready := FALSE;
FSteps[10].Children[2].Complete := TRUE;
FSteps[10].Children[2].Result := E_Result.Passed;
FSteps[10].Children[3].State := E_State.Completed;
FSteps[10].Children[3].Ready := FALSE;
FSteps[10].Children[3].Complete := TRUE;
FSteps[10].Children[3].Result := E_Result.Passed;
FSteps[10].ExpectedFinished := TRUE;
FSteps[10].MaxActiveChildCount := 0;
{endregion}
END_METHOD

END_FUNCTION_BLOCK

// ---- SelfTests/TestCases/TestSuite_ParallelSlotsOrchestration/Test_SlotsFirstFittingAdmission.TcPOU
{region 'Documentation'}
(*!
<summary>Selects fitting children only within the active slot and never bypasses a blocked group with a later-slot Start.</summary>
<description>
Child 1 waits for capacity while child 2 in the same slot fits and completes.
Child 3 always fits but belongs to slot 2, so even an otherwise idle slot 1 must wait
for child 1. Reservation responses isolate selection from Event Buffer arithmetic.
</description>
*)
{endregion}
FUNCTION_BLOCK Test_SlotsFirstFittingAdmission EXTENDS OrchestrationTestBase

SUPER^();

{region 'Documentation'}
(*!
<summary>Defines slot-group stimuli and per-cycle dispatch, completion and reservation expectations.</summary>
*)
{endregion}
METHOD PROTECTED ConfigureScenario
FChildSlots[1] := 1;
FChildSlots[2] := 1;
FChildSlots[3] := 2;
FStepCount := 10;

{region "01 - Observe initial readiness"}
FSteps[1].Task := E_OrchestratorTask.Idle;
FSteps[1].ExpectedReady := TRUE;
FSteps[1].MaxActiveChildCount := 0;
{endregion}

{region "02 - Skip blocked child 1 and start same-slot child 2"}
FSteps[2].Children[2].State := E_State.Running;
FSteps[2].Children[2].Ready := FALSE;
FSteps[2].ExecutionReservationResults[1] := E_EventReservationResult.WaitingForCapacity;
FSteps[2].ExpectedUnacceptedExecutionReservations[1] := 1;
FSteps[2].ExpectedStartChild := 2;
FSteps[2].ExpectedSlot := 1;
FSteps[2].ExpectedReservations[2] := 1;
FSteps[2].MaxActiveChildCount := 1;
{endregion}

{region "03 - Child 2 completes while child 1 still waits"}
FSteps[3].Children[2].State := E_State.Completed;
FSteps[3].Children[2].Ready := FALSE;
FSteps[3].Children[2].Complete := TRUE;
FSteps[3].Children[2].Result := E_Result.Passed;
FSteps[3].ExecutionReservationResults[1] := E_EventReservationResult.WaitingForCapacity;
FSteps[3].ExpectedUnacceptedExecutionReservations[1] := 1;
FSteps[3].ExpectedSlot := 1;
FSteps[3].ExpectedReservations[2] := 1;
FSteps[3].MaxActiveChildCount := 1;
{endregion}

{region "04 - Release child 2 but do not try the fitting later-slot child"}
FSteps[4].Children[2].State := E_State.Completed;
FSteps[4].Children[2].Ready := FALSE;
FSteps[4].Children[2].Complete := TRUE;
FSteps[4].Children[2].Result := E_Result.Passed;
FSteps[4].ExecutionReservationResults[1] := E_EventReservationResult.WaitingForCapacity;
FSteps[4].ExpectedUnacceptedExecutionReservations[1] := 1;
FSteps[4].ExpectedSlot := 1;
FSteps[4].ExpectedReleasedEntries[2] := 1;
FSteps[4].MaxActiveChildCount := 0;
{endregion}

{region "05 - Admit child 1 when its reservation becomes available"}
FSteps[5].Children[1].State := E_State.Running;
FSteps[5].Children[1].Ready := FALSE;
FSteps[5].Children[2].State := E_State.Completed;
FSteps[5].Children[2].Ready := FALSE;
FSteps[5].Children[2].Complete := TRUE;
FSteps[5].Children[2].Result := E_Result.Passed;
FSteps[5].ExpectedStartChild := 1;
FSteps[5].ExpectedSlot := 1;
FSteps[5].ExpectedReservations[1] := 1;
FSteps[5].MaxActiveChildCount := 1;
{endregion}

{region "06 - Child 1 completes before any later-slot Start"}
FSteps[6].Children[1].State := E_State.Completed;
FSteps[6].Children[1].Ready := FALSE;
FSteps[6].Children[1].Complete := TRUE;
FSteps[6].Children[1].Result := E_Result.Passed;
FSteps[6].Children[2].State := E_State.Completed;
FSteps[6].Children[2].Ready := FALSE;
FSteps[6].Children[2].Complete := TRUE;
FSteps[6].Children[2].Result := E_Result.Passed;
FSteps[6].ExpectedSlot := 1;
FSteps[6].ExpectedReservations[1] := 1;
FSteps[6].MaxActiveChildCount := 1;
{endregion}

{region "07 - Release child 1 and select the next slot"}
FSteps[7].Children[1].State := E_State.Completed;
FSteps[7].Children[1].Ready := FALSE;
FSteps[7].Children[1].Complete := TRUE;
FSteps[7].Children[1].Result := E_Result.Passed;
FSteps[7].Children[2].State := E_State.Completed;
FSteps[7].Children[2].Ready := FALSE;
FSteps[7].Children[2].Complete := TRUE;
FSteps[7].Children[2].Result := E_Result.Passed;
FSteps[7].ExpectedSlot := 2;
FSteps[7].ExpectedReleasedEntries[1] := 1;
FSteps[7].MaxActiveChildCount := 0;
{endregion}

{region "08 - Start the previously excluded child which completes immediately"}
FSteps[8].Children[1].State := E_State.Completed;
FSteps[8].Children[1].Ready := FALSE;
FSteps[8].Children[1].Complete := TRUE;
FSteps[8].Children[1].Result := E_Result.Passed;
FSteps[8].Children[2].State := E_State.Completed;
FSteps[8].Children[2].Ready := FALSE;
FSteps[8].Children[2].Complete := TRUE;
FSteps[8].Children[2].Result := E_Result.Passed;
FSteps[8].Children[3].State := E_State.Completed;
FSteps[8].Children[3].Ready := FALSE;
FSteps[8].Children[3].Complete := TRUE;
FSteps[8].Children[3].Result := E_Result.Passed;
FSteps[8].ExpectedStartChild := 3;
FSteps[8].ExpectedSlot := 2;
FSteps[8].ExpectedReservations[3] := 1;
FSteps[8].MaxActiveChildCount := 1;
{endregion}

{region "09 - Confirm the final Start and release its reservation"}
FSteps[9].Children[1].State := E_State.Completed;
FSteps[9].Children[1].Ready := FALSE;
FSteps[9].Children[1].Complete := TRUE;
FSteps[9].Children[1].Result := E_Result.Passed;
FSteps[9].Children[2].State := E_State.Completed;
FSteps[9].Children[2].Ready := FALSE;
FSteps[9].Children[2].Complete := TRUE;
FSteps[9].Children[2].Result := E_Result.Passed;
FSteps[9].Children[3].State := E_State.Completed;
FSteps[9].Children[3].Ready := FALSE;
FSteps[9].Children[3].Complete := TRUE;
FSteps[9].Children[3].Result := E_Result.Passed;
FSteps[9].ExpectedFinished := TRUE;
FSteps[9].ExpectedReleasedEntries[3] := 1;
FSteps[9].MaxActiveChildCount := 0;
{endregion}

{region "10 - Keep final completion stable without repeating admission"}
FSteps[10].Children[1].State := E_State.Completed;
FSteps[10].Children[1].Ready := FALSE;
FSteps[10].Children[1].Complete := TRUE;
FSteps[10].Children[1].Result := E_Result.Passed;
FSteps[10].Children[2].State := E_State.Completed;
FSteps[10].Children[2].Ready := FALSE;
FSteps[10].Children[2].Complete := TRUE;
FSteps[10].Children[2].Result := E_Result.Passed;
FSteps[10].Children[3].State := E_State.Completed;
FSteps[10].Children[3].Ready := FALSE;
FSteps[10].Children[3].Complete := TRUE;
FSteps[10].Children[3].Result := E_Result.Passed;
FSteps[10].ExpectedFinished := TRUE;
FSteps[10].MaxActiveChildCount := 0;
{endregion}
END_METHOD

END_FUNCTION_BLOCK

// ---- SelfTests/TestCases/TestSuite_ParallelSlotsOrchestration/Test_SlotsMissingStartReaction.TcPOU
{region 'Documentation'}
(*!
<summary>Rejects a missing Start reaction at the first-slot boundary without starting the next slot.</summary>
<description>
Child 1 completes immediately. Child 2 is then admitted but remains Idle.
The pending Start must be rejected once, its reservation released and child 3 left
untouched in slot 2. Repeated calls must preserve the Error without repeating diagnostics.
</description>
*)
{endregion}
FUNCTION_BLOCK Test_SlotsMissingStartReaction EXTENDS OrchestrationTestBase

SUPER^();

{region 'Documentation'}
(*!
<summary>Defines boundary stimuli and expected child requests, reservation cleanup and isolated diagnostics.</summary>
*)
{endregion}
METHOD PROTECTED ConfigureScenario
FChildSlots[1] := 1;
FChildSlots[2] := 1;
FChildSlots[3] := 2;
FStepCount := 5;

{region "01 - Observe initial readiness"}
FSteps[1].Task := E_OrchestratorTask.Idle;
FSteps[1].ExpectedReady := TRUE;
FSteps[1].MaxActiveChildCount := 0;
{endregion}

{region "02 - Child 1 completes immediately after Start"}
FSteps[2].Children[1].State := E_State.Completed;
FSteps[2].Children[1].Ready := FALSE;
FSteps[2].Children[1].Complete := TRUE;
FSteps[2].Children[1].Result := E_Result.Passed;
FSteps[2].ExpectedStartChild := 1;
FSteps[2].ExpectedSlot := 1;
FSteps[2].ExpectedReservations[1] := 1;
FSteps[2].MaxActiveChildCount := 1;
{endregion}

{region "03 - Start child 2 but retain its Idle observation"}
FSteps[3].Children[1].State := E_State.Completed;
FSteps[3].Children[1].Ready := FALSE;
FSteps[3].Children[1].Complete := TRUE;
FSteps[3].Children[1].Result := E_Result.Passed;
FSteps[3].ExpectedStartChild := 2;
FSteps[3].ExpectedSlot := 1;
FSteps[3].ExpectedReservations[2] := 1;
FSteps[3].ExpectedReleasedEntries[1] := 1;
FSteps[3].MaxActiveChildCount := 1;
{endregion}

{region "04 - Reject the missing reaction and release the pending reservation"}
FSteps[4].Children[1].State := E_State.Completed;
FSteps[4].Children[1].Ready := FALSE;
FSteps[4].Children[1].Complete := TRUE;
FSteps[4].Children[1].Result := E_Result.Passed;
FSteps[4].ExpectedSlot := 1;
FSteps[4].ExpectedResult := E_Result.Error;
FSteps[4].ExpectedDiagnosticCount := 1;
FSteps[4].ExpectedReleasedEntries[2] := 1;
FSteps[4].MaxActiveChildCount := 0;
{endregion}

{region "05 - Keep the next slot blocked without repeating the diagnostic"}
FSteps[5].Children[1].State := E_State.Completed;
FSteps[5].Children[1].Ready := FALSE;
FSteps[5].Children[1].Complete := TRUE;
FSteps[5].Children[1].Result := E_Result.Passed;
FSteps[5].ExpectedSlot := 1;
FSteps[5].ExpectedResult := E_Result.Error;
FSteps[5].ExpectedDiagnosticCount := 1;
FSteps[5].MaxActiveChildCount := 0;
{endregion}
END_METHOD

END_FUNCTION_BLOCK

// ---- SelfTests/TestCases/TestSuite_ParallelSlotsOrchestration/Test_SlotsNextSlotReadinessLost.TcPOU
{region 'Documentation'}
(*!
<summary>Prevents dispatch when the next slot loses readiness after initially valid admission.</summary>
<description>
All children are initially ready. While slot 1 completes, child 3 loses its readiness.
Selecting slot 2 must not dispatch it; the next check reports the readiness failure.
Later readiness recovery must not clear the held Error or trigger a Start.
</description>
*)
{endregion}
FUNCTION_BLOCK Test_SlotsNextSlotReadinessLost EXTENDS OrchestrationTestBase

SUPER^();

{region 'Documentation'}
(*!
<summary>Defines boundary stimuli and expected child requests, reservation cleanup and isolated diagnostics.</summary>
*)
{endregion}
METHOD PROTECTED ConfigureScenario
FChildSlots[1] := 1;
FChildSlots[2] := 1;
FChildSlots[3] := 2;
FStepCount := 7;

{region "01 - Observe all children initially ready"}
FSteps[1].Task := E_OrchestratorTask.Idle;
FSteps[1].ExpectedReady := TRUE;
FSteps[1].MaxActiveChildCount := 0;
{endregion}

{region "02 - Start child 1 in slot 1"}
FSteps[2].Children[1].State := E_State.Running;
FSteps[2].Children[1].Ready := FALSE;
FSteps[2].ExpectedStartChild := 1;
FSteps[2].ExpectedSlot := 1;
FSteps[2].ExpectedReservations[1] := 1;
FSteps[2].MaxActiveChildCount := 1;
{endregion}

{region "03 - Start child 2 and complete slot 1 while child 3 loses readiness"}
FSteps[3].Children[1].State := E_State.Completed;
FSteps[3].Children[1].Ready := FALSE;
FSteps[3].Children[1].Complete := TRUE;
FSteps[3].Children[1].Result := E_Result.Passed;
FSteps[3].Children[2].State := E_State.Completed;
FSteps[3].Children[2].Ready := FALSE;
FSteps[3].Children[2].Complete := TRUE;
FSteps[3].Children[2].Result := E_Result.Passed;
FSteps[3].Children[3].Ready := FALSE;
FSteps[3].ExpectedStartChild := 2;
FSteps[3].ExpectedSlot := 1;
FSteps[3].ExpectedReservations[1] := 1;
FSteps[3].ExpectedReservations[2] := 1;
FSteps[3].MaxActiveChildCount := 2;
{endregion}

{region "04 - Release slot 1 and select slot 2 without dispatch"}
FSteps[4].Children[1].State := E_State.Completed;
FSteps[4].Children[1].Ready := FALSE;
FSteps[4].Children[1].Complete := TRUE;
FSteps[4].Children[1].Result := E_Result.Passed;
FSteps[4].Children[2].State := E_State.Completed;
FSteps[4].Children[2].Ready := FALSE;
FSteps[4].Children[2].Complete := TRUE;
FSteps[4].Children[2].Result := E_Result.Passed;
FSteps[4].Children[3].Ready := FALSE;
FSteps[4].ExpectedSlot := 2;
FSteps[4].ExpectedReleasedEntries[1] := 1;
FSteps[4].ExpectedReleasedEntries[2] := 1;
FSteps[4].MaxActiveChildCount := 0;
{endregion}

{region "05 - Reject the now unready next-slot child before Start"}
FSteps[5].Children[1].State := E_State.Completed;
FSteps[5].Children[1].Ready := FALSE;
FSteps[5].Children[1].Complete := TRUE;
FSteps[5].Children[1].Result := E_Result.Passed;
FSteps[5].Children[2].State := E_State.Completed;
FSteps[5].Children[2].Ready := FALSE;
FSteps[5].Children[2].Complete := TRUE;
FSteps[5].Children[2].Result := E_Result.Passed;
FSteps[5].Children[3].Ready := FALSE;
FSteps[5].ExpectedSlot := 2;
FSteps[5].ExpectedResult := E_Result.Error;
FSteps[5].ExpectedDiagnosticCount := 1;
FSteps[5].MaxActiveChildCount := 0;
{endregion}

{region "06 - Restore readiness without clearing the held Error"}
FSteps[6].Children[1].State := E_State.Completed;
FSteps[6].Children[1].Ready := FALSE;
FSteps[6].Children[1].Complete := TRUE;
FSteps[6].Children[1].Result := E_Result.Passed;
FSteps[6].Children[2].State := E_State.Completed;
FSteps[6].Children[2].Ready := FALSE;
FSteps[6].Children[2].Complete := TRUE;
FSteps[6].Children[2].Result := E_Result.Passed;
FSteps[6].ExpectedSlot := 2;
FSteps[6].ExpectedResult := E_Result.Error;
FSteps[6].ExpectedDiagnosticCount := 1;
FSteps[6].MaxActiveChildCount := 0;
{endregion}

{region "07 - Do not resume dispatch after readiness recovery"}
FSteps[7].Children[1].State := E_State.Completed;
FSteps[7].Children[1].Ready := FALSE;
FSteps[7].Children[1].Complete := TRUE;
FSteps[7].Children[1].Result := E_Result.Passed;
FSteps[7].Children[2].State := E_State.Completed;
FSteps[7].Children[2].Ready := FALSE;
FSteps[7].Children[2].Complete := TRUE;
FSteps[7].Children[2].Result := E_Result.Passed;
FSteps[7].ExpectedSlot := 2;
FSteps[7].ExpectedResult := E_Result.Error;
FSteps[7].ExpectedDiagnosticCount := 1;
FSteps[7].MaxActiveChildCount := 0;
{endregion}
END_METHOD

END_FUNCTION_BLOCK

// ---- SelfTests/TestCases/TestSuite_ParallelSlotsOrchestration/Test_SlotsAbortAtBoundary.TcPOU
{region 'Documentation'}
(*!
<summary>Accepts an immediately completed pending Start when Abort replaces execution at the slot boundary.</summary>
<description>
Both children in slot 1 complete directly after their respective Start requests.
Before the second Start is confirmed, the owner selects Abort. Confirmation and
reservation cleanup must finish without starting child 3 or aborting already stopped children.
</description>
*)
{endregion}
FUNCTION_BLOCK Test_SlotsAbortAtBoundary EXTENDS OrchestrationTestBase

SUPER^();

{region 'Documentation'}
(*!
<summary>Defines boundary stimuli and expected child requests, reservation cleanup and isolated diagnostics.</summary>
*)
{endregion}
METHOD PROTECTED ConfigureScenario
FChildSlots[1] := 1;
FChildSlots[2] := 1;
FChildSlots[3] := 2;
FStepCount := 5;

{region "01 - Observe initial readiness"}
FSteps[1].Task := E_OrchestratorTask.Idle;
FSteps[1].ExpectedReady := TRUE;
FSteps[1].MaxActiveChildCount := 0;
{endregion}

{region "02 - Child 1 completes immediately after Start"}
FSteps[2].Children[1].State := E_State.Completed;
FSteps[2].Children[1].Ready := FALSE;
FSteps[2].Children[1].Complete := TRUE;
FSteps[2].Children[1].Result := E_Result.Passed;
FSteps[2].ExpectedStartChild := 1;
FSteps[2].ExpectedSlot := 1;
FSteps[2].ExpectedReservations[1] := 1;
FSteps[2].MaxActiveChildCount := 1;
{endregion}

{region "03 - Child 2 completes immediately with Start confirmation pending"}
FSteps[3].Children[1].State := E_State.Completed;
FSteps[3].Children[1].Ready := FALSE;
FSteps[3].Children[1].Complete := TRUE;
FSteps[3].Children[1].Result := E_Result.Passed;
FSteps[3].Children[2].State := E_State.Completed;
FSteps[3].Children[2].Ready := FALSE;
FSteps[3].Children[2].Complete := TRUE;
FSteps[3].Children[2].Result := E_Result.Passed;
FSteps[3].ExpectedStartChild := 2;
FSteps[3].ExpectedSlot := 1;
FSteps[3].ExpectedReservations[2] := 1;
FSteps[3].ExpectedReleasedEntries[1] := 1;
FSteps[3].MaxActiveChildCount := 1;
{endregion}

{region "04 - Abort confirms completion and releases the pending reservation"}
FSteps[4].Task := E_OrchestratorTask.Abort;
FSteps[4].Children[1].State := E_State.Completed;
FSteps[4].Children[1].Ready := FALSE;
FSteps[4].Children[1].Complete := TRUE;
FSteps[4].Children[1].Result := E_Result.Passed;
FSteps[4].Children[2].State := E_State.Completed;
FSteps[4].Children[2].Ready := FALSE;
FSteps[4].Children[2].Complete := TRUE;
FSteps[4].Children[2].Result := E_Result.Passed;
FSteps[4].ExpectedAbortFinished := TRUE;
FSteps[4].ExpectedReleasedEntries[2] := 1;
FSteps[4].MaxActiveChildCount := 0;
{endregion}

{region "05 - Keep Abort complete without starting the next slot"}
FSteps[5].Task := E_OrchestratorTask.Abort;
FSteps[5].Children[1].State := E_State.Completed;
FSteps[5].Children[1].Ready := FALSE;
FSteps[5].Children[1].Complete := TRUE;
FSteps[5].Children[1].Result := E_Result.Passed;
FSteps[5].Children[2].State := E_State.Completed;
FSteps[5].Children[2].Ready := FALSE;
FSteps[5].Children[2].Complete := TRUE;
FSteps[5].Children[2].Result := E_Result.Passed;
FSteps[5].ExpectedAbortFinished := TRUE;
FSteps[5].MaxActiveChildCount := 0;
{endregion}
END_METHOD

END_FUNCTION_BLOCK

// ---- SelfTests/TestSuites/TestSuite_TestSuiteConfigurationBuilder.TcPOU
{region 'Documentation'}
(*!
<summary>Checks the Test Suite builder directly without executing registered child lifecycles.</summary>
*)
{endregion}
FUNCTION_BLOCK TestSuite_TestSuiteConfigurationBuilder EXTENDS TestSuiteBase
VAR
    FSerial : Test_SuiteBuilderSerial;
    FParallel : Test_SuiteBuilderParallel;
    FSlotInsertion : Test_SuiteBuilderSlotInsertion;
    FCapacity : Test_SuiteBuilderCapacity;
    FRegistrationErrors : Test_SuiteBuilderRegistrationErrors;
    FFinalizeReuse : Test_SuiteBuilderFinalizeReuse;
    FTestCases : ARRAY[1..TestCaseCapacity] OF I_TestCase;
END_VAR
VAR CONSTANT
    TestCaseCapacity : UINT := 6;
END_VAR

SUPER^();

{region 'Documentation'}
(*!
<summary>Initializes and registers the six independent builder scenarios for serial execution.</summary>
*)
{endregion}
METHOD PROTECTED Configure
VAR_IN_OUT
    // SA0167: Borrowed owner builder; no temporary instance is created.
    {attribute 'analysis' := '-167'}
    Builder : TestSuiteConfigurationBuilder; //! Borrowed owner configuration builder used only during this Configure call; register this owner's concrete children.
END_VAR
VAR
    TestConfig : ST_TestCaseConfig;
END_VAR
Builder.Initialize(Mode := E_OrchestrationMode.Serial,
    TestCases := FTestCases);

FSerial.Initialize(Parent := THIS^,
    TestName := 'Serial',
    Config := TestConfig);
Builder.Register(TestCase := FSerial);

FParallel.Initialize(Parent := THIS^,
    TestName := 'Parallel',
    Config := TestConfig);
Builder.Register(TestCase := FParallel);

FSlotInsertion.Initialize(Parent := THIS^,
    TestName := 'SlotInsertion',
    Config := TestConfig);
Builder.Register(TestCase := FSlotInsertion);

FCapacity.Initialize(Parent := THIS^,
    TestName := 'Capacity',
    Config := TestConfig);
Builder.Register(TestCase := FCapacity);

FRegistrationErrors.Initialize(Parent := THIS^,
    TestName := 'RegistrationErrors',
    Config := TestConfig);
Builder.Register(TestCase := FRegistrationErrors);

FFinalizeReuse.Initialize(Parent := THIS^,
    TestName := 'FinalizeReuse',
    Config := TestConfig);
Builder.Register(TestCase := FFinalizeReuse);
END_METHOD

{region 'Documentation'}
(*!
<summary>Returns a registered scenario using the actual array index.</summary>
*)
{endregion}
METHOD PUBLIC GetTestCase : I_TestCase //! Typed child interface at the original array index; zero when no entry is available.
VAR_INPUT
    Index : DINT; //! Original occupied child-array index, rather than an ordinal position.
END_VAR
GetTestCase := 0;
IF (ChildCount = 0) OR (Index < ChildArrayLowerBound)
    OR (DINT_TO_LINT(Index) >= DINT_TO_LINT(ChildArrayLowerBound) + UINT_TO_LINT(ChildCount)) THEN
    RETURN;
END_IF;

GetTestCase := FTestCases[Index];
END_METHOD

{region 'Documentation'}
(*!
<summary>Calls the six owned scenarios once per initialized Suite cycle.</summary>
*)
{endregion}
METHOD PROTECTED ProcessTestCases
FSerial();
FParallel();
FSlotInsertion();
FCapacity();
FRegistrationErrors();
FFinalizeReuse();
END_METHOD

END_FUNCTION_BLOCK

// ---- SelfTests/TestCases/TestSuite_TestSuiteConfigurationBuilder/Test_SuiteBuilderSerial.TcPOU
{region 'Documentation'}
(*!
<summary>Checks Serial registration with shifted bounds and unused capacity.</summary>
<description>Child mocks are inert interface identities and slot storage only; no child initialization or FB call is performed.</description>
*)
{endregion}
FUNCTION_BLOCK Test_SuiteBuilderSerial EXTENDS TestCaseBase
VAR
    FBuilder : TestSuiteConfigurationBuilder;
    FCases : ARRAY[4..7] OF I_TestCase;
    FChildA : TestCaseMock;
    FChildB : TestCaseMock;
    FChildC : TestCaseMock;
    FScenarioExecuted : BOOL;
    FChecksEvaluated : BOOL;
    FClearing : AssertTrue;
    FClearingMatches : BOOL;
    FRegistration : AssertTrue;
    FRegistrationMatches : BOOL;
    FOrder : AssertTrue;
    FOrderMatches : BOOL;
    FSlots : AssertTrue;
    FSlotsMatches : BOOL;
    FMetadata : AssertTrue;
    FMetadataMatches : BOOL;
    FFinalization : AssertTrue;
    FFinalizationMatches : BOOL;
END_VAR

SUPER^();

{region 'Documentation'}
(*!
<summary>Contributes each owned Assertion once without executing it.</summary>
*)
{endregion}
METHOD PROTECTED AggregateResults
VAR_INPUT
    Aggregator : I_ResultAggregator; //! Borrowed result sink owned by the outer Test Case; add this test's checking Assertions without resetting or retaining the sink.
END_VAR
Aggregator.AddProvider(Provider := FClearing);
Aggregator.AddProvider(Provider := FRegistration);
Aggregator.AddProvider(Provider := FOrder);
Aggregator.AddProvider(Provider := FSlots);
Aggregator.AddProvider(Provider := FMetadata);
Aggregator.AddProvider(Provider := FFinalization);
END_METHOD

{region 'Documentation'}
(*!
<summary>Requires successful base and owned Assertion initialization.</summary>
*)
{endregion}
METHOD PROTECTED CheckInitialization : BOOL //! TRUE when the inherited initialization check and this concrete fixture check both accept the setup.
CheckInitialization := FALSE;
IF NOT SUPER^.CheckInitialization() THEN
    RETURN;
END_IF;

CheckInitialization := FClearing.IsInitialized
    AND FRegistration.IsInitialized
    AND FOrder.IsInitialized
    AND FSlots.IsInitialized
    AND FMetadata.IsInitialized
    AND FFinalization.IsInitialized;
END_METHOD

{region 'Documentation'}
(*!
<summary>Configures one direct builder scenario and its named Assertions.</summary>
*)
{endregion}
METHOD PROTECTED Configure
FPreparationStateCount := 0;
FTestStateCount := 1;
FScenarioExecuted := FALSE;
FChecksEvaluated := FALSE;

FClearingMatches := FALSE;
FClearing.Initialize(Parent := THIS^,
    AssertionName := 'Clearing');
FRegistrationMatches := FALSE;
FRegistration.Initialize(Parent := THIS^,
    AssertionName := 'Registration');
FOrderMatches := FALSE;
FOrder.Initialize(Parent := THIS^,
    AssertionName := 'Order');
FSlotsMatches := FALSE;
FSlots.Initialize(Parent := THIS^,
    AssertionName := 'Slots');
FMetadataMatches := FALSE;
FMetadata.Initialize(Parent := THIS^,
    AssertionName := 'Metadata');
FFinalizationMatches := FALSE;
FFinalization.Initialize(Parent := THIS^,
    AssertionName := 'Finalization');
END_METHOD

{region 'Documentation'}
(*!
<summary>Completes Abort immediately; no asynchronous resource operation is started.</summary>
*)
{endregion}
METHOD PROTECTED ProcessAbort
VAR_INPUT
    Enable : BOOL; //! Phase permission supplied by the owning Test Case; FALSE does not authorize progression, while observation may continue.
END_VAR
IF Enable THEN
    CompleteAbort();
END_IF;
END_METHOD

{region 'Documentation'}
(*!
<summary>Evaluates recorded observations and consumes pending resets on disabled calls.</summary>
*)
{endregion}
METHOD PROTECTED ProcessAssertions
VAR_INPUT
    Enable : BOOL; //! Phase permission supplied by the owning Test Case; FALSE does not authorize progression, while observation may continue.
END_VAR
FClearing(Enable := Enable,
    State := State,
    IN := FClearingMatches);

FRegistration(Enable := Enable,
    State := State,
    IN := FRegistrationMatches);

FOrder(Enable := Enable,
    State := State,
    IN := FOrderMatches);

FSlots(Enable := Enable,
    State := State,
    IN := FSlotsMatches);

FMetadata(Enable := Enable,
    State := State,
    IN := FMetadataMatches);

FFinalization(Enable := Enable,
    State := State,
    IN := FFinalizationMatches);

IF Enable AND FClearing.EvaluationActive
    AND FRegistration.EvaluationActive
    AND FOrder.EvaluationActive
    AND FSlots.EvaluationActive
    AND FMetadata.EvaluationActive
    AND FFinalization.EvaluationActive THEN
    FChecksEvaluated := TRUE;
END_IF;
END_METHOD

{region 'Documentation'}
(*!
<summary>No Preparation phase is needed for synchronous builder calls.</summary>
*)
{endregion}
METHOD PROTECTED ProcessPreparations
VAR_INPUT
    // SA0033: Required override signature; this scenario has no Preparation work.
    {attribute 'analysis' := '-33'}
    Enable : BOOL; //! Phase permission supplied by the owning Test Case; FALSE does not authorize progression, while observation may continue.
END_VAR
END_METHOD

{region 'Documentation'}
(*!
<summary>Clears recorded checks and Assertion results; each scenario initializes its own builder.</summary>
*)
{endregion}
METHOD PROTECTED ProcessReset
FScenarioExecuted := FALSE;
FChecksEvaluated := FALSE;
FClearingMatches := FALSE;
FClearing.Reset();
FRegistrationMatches := FALSE;
FRegistration.Reset();
FOrderMatches := FALSE;
FOrder.Reset();
FSlotsMatches := FALSE;
FSlots.Reset();
FMetadataMatches := FALSE;
FMetadata.Reset();
FFinalizationMatches := FALSE;
FFinalization.Reset();
CompleteReset();
END_METHOD

{region 'Documentation'}
(*!
<summary>Runs setup operations once, then completes after their observations have been evaluated.</summary>
*)
{endregion}
METHOD PROTECTED ProcessTests
VAR_INPUT
    Enable : BOOL; //! Phase permission supplied by the owning Test Case; FALSE does not authorize progression, while observation may continue.
END_VAR
IF NOT Enable THEN
    RETURN;
END_IF;

IF FChecksEvaluated THEN
    CompleteTests();
ELSIF NOT FScenarioExecuted THEN
    RunScenario();
    FScenarioExecuted := TRUE;
END_IF;
END_METHOD

{region 'Documentation'}
(*!
<summary>Checks Serial registration with shifted bounds and unused capacity.</summary>
*)
{endregion}
METHOD PRIVATE RunScenario
VAR
    ChildA : I_TestCase;
    ChildB : I_TestCase;
    ChildC : I_TestCase;
    AcceptedA : BOOL;
    AcceptedB : BOOL;
    AcceptedC : BOOL;
    Config : ST_TestCaseCollectionConfig;
END_VAR
ChildA := FChildA;
ChildB := FChildB;
ChildC := FChildC;
FCases[4] := ChildA;
FCases[5] := ChildB;
FCases[6] := ChildC;
FCases[7] := ChildA;
FBuilder.Initialize(Mode := E_OrchestrationMode.Serial,
    TestCases := FCases);
FClearingMatches := (FCases[4] = 0) AND (FCases[5] = 0)
    AND (FCases[6] = 0) AND (FCases[7] = 0)
    AND (FBuilder.Count = 0) AND NOT FBuilder.IsValid AND NOT FBuilder.IsFinalized;

AcceptedA := FBuilder.Register(TestCase := ChildC);
AcceptedB := FBuilder.Register(TestCase := ChildA);
AcceptedC := FBuilder.Register(TestCase := ChildB);
FRegistrationMatches := AcceptedA AND AcceptedB AND AcceptedC;
FOrderMatches := (FCases[4] = ChildC) AND (FCases[5] = ChildA)
    AND (FCases[6] = ChildB) AND (FCases[7] = 0);
FSlotsMatches := (FChildC.ExecutionSlot = 1) AND (FChildA.ExecutionSlot = 2)
    AND (FChildB.ExecutionSlot = 3);
FMetadataMatches := (FBuilder.FirstIndex = 4) AND (FBuilder.LastIndex = 7)
    AND (FBuilder.Count = 3) AND (FBuilder.Mode = E_OrchestrationMode.Serial);

Config := FBuilder.Finalize();
FFinalizationMatches := Config.IsValid AND FBuilder.IsValid AND FBuilder.IsFinalized
    AND (Config.FirstIndex = 4) AND (Config.LastIndex = 7) AND (Config.Count = 3)
    AND (Config.Mode = E_OrchestrationMode.Serial);
END_METHOD

END_FUNCTION_BLOCK

// ---- Framework/TestCases/POU/TestCaseMock.TcPOU
{region 'Documentation'}
(*!
<summary>Simple Test Case double using the real base lifecycle and one simulated Assertion
result.</summary>
<description>
No Preparation or concrete Assertion instances are owned. Initialize through the inherited
API; Ready gates Start and Completed plus MinimumTestDuration gate normal completion.

MinimumTestDuration defaults to T#100ms and survives Initialize and Reset. Error, Abort and
owner timeout are not delayed. ResultValue contributes one counted result; this is a lifecycle
double, not evidence from real Assertions.
</description>
*)
{endregion}
FUNCTION_BLOCK TestCaseMock EXTENDS TestCaseBase
VAR_INPUT
    Ready : BOOL := TRUE; //! Application readiness gate for starting the mock; default TRUE.
    Completed : BOOL := TRUE; //! Allows normal mock completion after MinimumTestDuration; default TRUE.
    ResultValue : E_Result := E_Result.Passed; //! Simulated test outcome; default Passed. Lifecycle errors can still escalate the owner result.
END_VAR
VAR
    FMinimumTestDuration : TIME := T#100ms;
END_VAR

SUPER^();

{region 'Documentation'}
(*!
<summary>Contributes one simulated Assertion result.</summary>
<description>
Contributes NotEvaluated in Reset and Idle, otherwise ResultValue, including during Completed.
The base retains its completed owner result independently of the refreshed counter snapshot.
</description>
*)
{endregion}
METHOD PROTECTED AggregateResults
VAR_INPUT
    Aggregator : I_ResultAggregator; //! Owner-held contribution interface; add each child once without resetting or retaining this interface.
END_VAR
IF IsResetting OR (State = E_State.Idle) THEN
    Aggregator.AddResult(Result := E_Result.NotEvaluated);
    RETURN;
END_IF;
Aggregator.AddResult(Result := ResultValue);
END_METHOD

{region 'Documentation'}
(*!
<summary>Configures no Preparation phase and one Test state; retains caller settings.</summary>
*)
{endregion}
METHOD PROTECTED Configure
FPreparationStateCount := 0;
FTestStateCount := 1;
END_METHOD

{region 'Documentation'}
(*!
<summary>Combines base prerequisites with the externally controlled ready release.</summary>
*)
{endregion}
{attribute 'monitoring' := 'call'}
PROPERTY PUBLIC IsReady : BOOL //! Combines base prerequisites with the externally controlled ready release.
GET // PUBLIC
IsReady := SUPER^.IsReady AND Ready;
END_GET
END_PROPERTY

{region 'Documentation'}
(*!
<summary>Minimum duration of the Test phase; zero permits immediate normal completion.</summary>
<description>
Does not delay Abort, Error or the owner timeout. Initialize and Reset retain this
setting.
</description>
*)
{endregion}
{attribute 'monitoring' := 'call'}
PROPERTY PUBLIC MinimumTestDuration : TIME //! Minimum duration of the Test phase; zero permits immediate normal completion.
GET // PUBLIC
MinimumTestDuration := FMinimumTestDuration;
END_GET
SET // PUBLIC
FMinimumTestDuration := MinimumTestDuration;
END_SET
END_PROPERTY

{region 'Documentation'}
(*!
<summary>Immediately completes the base-selected Abort/Error path when enabled.</summary>
*)
{endregion}
METHOD PROTECTED ProcessAbort
VAR_INPUT
    Enable : BOOL; //! TRUE while this hook's lifecycle phase is active; FALSE must not advance that phase.
END_VAR
IF Enable THEN
    CompleteAbort();
END_IF;
END_METHOD

{region 'Documentation'}
(*!
<summary>Intentionally executes no Assertions; AggregateResults supplies the injected child
outcome.</summary>
*)
{endregion}
METHOD PROTECTED ProcessAssertions
VAR_INPUT
    // SA0033: Required inherited hook; this mock owns no children for this phase.
    {attribute 'analysis' := '-33'}
    Enable : BOOL; //! TRUE while this hook's lifecycle phase is active; FALSE must not advance that phase.
END_VAR
RETURN;
END_METHOD

{region 'Documentation'}
(*!
<summary>No Preparations are owned or executed.</summary>
*)
{endregion}
METHOD PROTECTED ProcessPreparations
VAR_INPUT
    // SA0033: Required inherited hook; this mock owns no children for this phase.
    {attribute 'analysis' := '-33'}
    Enable : BOOL; //! TRUE while this hook's lifecycle phase is active; FALSE must not advance that phase.
END_VAR
RETURN;
END_METHOD

{region 'Documentation'}
(*!
<summary>Completes Reset immediately; base-owned state is reset by the base.</summary>
*)
{endregion}
METHOD PROTECTED ProcessReset
CompleteReset();
END_METHOD

{region 'Documentation'}
(*!
<summary>Completes the enabled Test phase when released and its minimum duration has
elapsed.</summary>
*)
{endregion}
METHOD PROTECTED ProcessTests
VAR_INPUT
    Enable : BOOL; //! TRUE while this hook's lifecycle phase is active; FALSE must not advance that phase.
END_VAR
IF NOT Enable THEN
    RETURN;
END_IF;

IF Completed AND (FStateTimer.ElapsedLTime >= TIME_TO_LTIME(FMinimumTestDuration)) THEN
    CompleteTests();
END_IF;
END_METHOD

END_FUNCTION_BLOCK

// ---- SelfTests/TestCases/TestSuite_TestSuiteConfigurationBuilder/Test_SuiteBuilderParallel.TcPOU
{region 'Documentation'}
(*!
<summary>Checks Parallel registration order and shared slot across negative array bounds.</summary>
<description>Child mocks are inert interface identities and slot storage only; no child initialization or FB call is performed.</description>
*)
{endregion}
FUNCTION_BLOCK Test_SuiteBuilderParallel EXTENDS TestCaseBase
VAR
    FBuilder : TestSuiteConfigurationBuilder;
    FCases : ARRAY[-2..1] OF I_TestCase;
    FChildA : TestCaseMock;
    FChildB : TestCaseMock;
    FScenarioExecuted : BOOL;
    FChecksEvaluated : BOOL;
    FRegistration : AssertTrue;
    FRegistrationMatches : BOOL;
    FOrder : AssertTrue;
    FOrderMatches : BOOL;
    FSlots : AssertTrue;
    FSlotsMatches : BOOL;
    FMetadata : AssertTrue;
    FMetadataMatches : BOOL;
    FFinalization : AssertTrue;
    FFinalizationMatches : BOOL;
END_VAR

SUPER^();

{region 'Documentation'}
(*!
<summary>Contributes each owned Assertion once without executing it.</summary>
*)
{endregion}
METHOD PROTECTED AggregateResults
VAR_INPUT
    Aggregator : I_ResultAggregator; //! Borrowed result sink owned by the outer Test Case; add this test's checking Assertions without resetting or retaining the sink.
END_VAR
Aggregator.AddProvider(Provider := FRegistration);
Aggregator.AddProvider(Provider := FOrder);
Aggregator.AddProvider(Provider := FSlots);
Aggregator.AddProvider(Provider := FMetadata);
Aggregator.AddProvider(Provider := FFinalization);
END_METHOD

{region 'Documentation'}
(*!
<summary>Requires successful base and owned Assertion initialization.</summary>
*)
{endregion}
METHOD PROTECTED CheckInitialization : BOOL //! TRUE when the inherited initialization check and this concrete fixture check both accept the setup.
CheckInitialization := FALSE;
IF NOT SUPER^.CheckInitialization() THEN
    RETURN;
END_IF;

CheckInitialization := FRegistration.IsInitialized
    AND FOrder.IsInitialized
    AND FSlots.IsInitialized
    AND FMetadata.IsInitialized
    AND FFinalization.IsInitialized;
END_METHOD

{region 'Documentation'}
(*!
<summary>Configures one direct builder scenario and its named Assertions.</summary>
*)
{endregion}
METHOD PROTECTED Configure
FPreparationStateCount := 0;
FTestStateCount := 1;
FScenarioExecuted := FALSE;
FChecksEvaluated := FALSE;

FRegistrationMatches := FALSE;
FRegistration.Initialize(Parent := THIS^,
    AssertionName := 'Registration');
FOrderMatches := FALSE;
FOrder.Initialize(Parent := THIS^,
    AssertionName := 'Order');
FSlotsMatches := FALSE;
FSlots.Initialize(Parent := THIS^,
    AssertionName := 'Slots');
FMetadataMatches := FALSE;
FMetadata.Initialize(Parent := THIS^,
    AssertionName := 'Metadata');
FFinalizationMatches := FALSE;
FFinalization.Initialize(Parent := THIS^,
    AssertionName := 'Finalization');
END_METHOD

{region 'Documentation'}
(*!
<summary>Completes Abort immediately; no asynchronous resource operation is started.</summary>
*)
{endregion}
METHOD PROTECTED ProcessAbort
VAR_INPUT
    Enable : BOOL; //! Phase permission supplied by the owning Test Case; FALSE does not authorize progression, while observation may continue.
END_VAR
IF Enable THEN
    CompleteAbort();
END_IF;
END_METHOD

{region 'Documentation'}
(*!
<summary>Evaluates recorded observations and consumes pending resets on disabled calls.</summary>
*)
{endregion}
METHOD PROTECTED ProcessAssertions
VAR_INPUT
    Enable : BOOL; //! Phase permission supplied by the owning Test Case; FALSE does not authorize progression, while observation may continue.
END_VAR
FRegistration(Enable := Enable,
    State := State,
    IN := FRegistrationMatches);

FOrder(Enable := Enable,
    State := State,
    IN := FOrderMatches);

FSlots(Enable := Enable,
    State := State,
    IN := FSlotsMatches);

FMetadata(Enable := Enable,
    State := State,
    IN := FMetadataMatches);

FFinalization(Enable := Enable,
    State := State,
    IN := FFinalizationMatches);

IF Enable AND FRegistration.EvaluationActive
    AND FOrder.EvaluationActive
    AND FSlots.EvaluationActive
    AND FMetadata.EvaluationActive
    AND FFinalization.EvaluationActive THEN
    FChecksEvaluated := TRUE;
END_IF;
END_METHOD

{region 'Documentation'}
(*!
<summary>No Preparation phase is needed for synchronous builder calls.</summary>
*)
{endregion}
METHOD PROTECTED ProcessPreparations
VAR_INPUT
    // SA0033: Required override signature; this scenario has no Preparation work.
    {attribute 'analysis' := '-33'}
    Enable : BOOL; //! Phase permission supplied by the owning Test Case; FALSE does not authorize progression, while observation may continue.
END_VAR
END_METHOD

{region 'Documentation'}
(*!
<summary>Clears recorded checks and Assertion results; each scenario initializes its own builder.</summary>
*)
{endregion}
METHOD PROTECTED ProcessReset
FScenarioExecuted := FALSE;
FChecksEvaluated := FALSE;
FRegistrationMatches := FALSE;
FRegistration.Reset();
FOrderMatches := FALSE;
FOrder.Reset();
FSlotsMatches := FALSE;
FSlots.Reset();
FMetadataMatches := FALSE;
FMetadata.Reset();
FFinalizationMatches := FALSE;
FFinalization.Reset();
CompleteReset();
END_METHOD

{region 'Documentation'}
(*!
<summary>Runs setup operations once, then completes after their observations have been evaluated.</summary>
*)
{endregion}
METHOD PROTECTED ProcessTests
VAR_INPUT
    Enable : BOOL; //! Phase permission supplied by the owning Test Case; FALSE does not authorize progression, while observation may continue.
END_VAR
IF NOT Enable THEN
    RETURN;
END_IF;

IF FChecksEvaluated THEN
    CompleteTests();
ELSIF NOT FScenarioExecuted THEN
    RunScenario();
    FScenarioExecuted := TRUE;
END_IF;
END_METHOD

{region 'Documentation'}
(*!
<summary>Checks Parallel registration order and shared slot across negative array bounds.</summary>
*)
{endregion}
METHOD PRIVATE RunScenario
VAR
    ChildA : I_TestCase;
    ChildB : I_TestCase;
    AcceptedA : BOOL;
    AcceptedB : BOOL;
    Config : ST_TestCaseCollectionConfig;
END_VAR
ChildA := FChildA;
ChildB := FChildB;
FBuilder.Initialize(Mode := E_OrchestrationMode.Parallel,
    TestCases := FCases);
AcceptedA := FBuilder.Register(TestCase := ChildB);
AcceptedB := FBuilder.Register(TestCase := ChildA);
FRegistrationMatches := AcceptedA AND AcceptedB;
FOrderMatches := (FCases[-2] = ChildB) AND (FCases[-1] = ChildA)
    AND (FCases[0] = 0) AND (FCases[1] = 0);
FSlotsMatches := (FChildA.ExecutionSlot = 1) AND (FChildB.ExecutionSlot = 1);
FMetadataMatches := (FBuilder.FirstIndex = -2) AND (FBuilder.LastIndex = 1)
    AND (FBuilder.Count = 2) AND (FBuilder.Mode = E_OrchestrationMode.Parallel);

Config := FBuilder.Finalize();
FFinalizationMatches := Config.IsValid AND FBuilder.IsValid AND FBuilder.IsFinalized
    AND (Config.FirstIndex = -2) AND (Config.LastIndex = 1) AND (Config.Count = 2)
    AND (Config.Mode = E_OrchestrationMode.Parallel);
END_METHOD

END_FUNCTION_BLOCK

// ---- SelfTests/TestCases/TestSuite_TestSuiteConfigurationBuilder/Test_SuiteBuilderSlotInsertion.TcPOU
{region 'Documentation'}
(*!
<summary>Checks stable insertion into two slots, including a temporary gap before Finalize.</summary>
<description>Child mocks are inert interface identities and slot storage only; no child initialization or FB call is performed.</description>
*)
{endregion}
FUNCTION_BLOCK Test_SuiteBuilderSlotInsertion EXTENDS TestCaseBase
VAR
    FBuilder : TestSuiteConfigurationBuilder;
    FCases : ARRAY[1..4] OF I_TestCase;
    FChildA : TestCaseMock;
    FChildB : TestCaseMock;
    FChildC : TestCaseMock;
    FChildD : TestCaseMock;
    FScenarioExecuted : BOOL;
    FChecksEvaluated : BOOL;
    FRegistration : AssertTrue;
    FRegistrationMatches : BOOL;
    FOrder : AssertTrue;
    FOrderMatches : BOOL;
    FSlots : AssertTrue;
    FSlotsMatches : BOOL;
    FFinalization : AssertTrue;
    FFinalizationMatches : BOOL;
END_VAR

SUPER^();

{region 'Documentation'}
(*!
<summary>Contributes each owned Assertion once without executing it.</summary>
*)
{endregion}
METHOD PROTECTED AggregateResults
VAR_INPUT
    Aggregator : I_ResultAggregator; //! Borrowed result sink owned by the outer Test Case; add this test's checking Assertions without resetting or retaining the sink.
END_VAR
Aggregator.AddProvider(Provider := FRegistration);
Aggregator.AddProvider(Provider := FOrder);
Aggregator.AddProvider(Provider := FSlots);
Aggregator.AddProvider(Provider := FFinalization);
END_METHOD

{region 'Documentation'}
(*!
<summary>Requires successful base and owned Assertion initialization.</summary>
*)
{endregion}
METHOD PROTECTED CheckInitialization : BOOL //! TRUE when the inherited initialization check and this concrete fixture check both accept the setup.
CheckInitialization := FALSE;
IF NOT SUPER^.CheckInitialization() THEN
    RETURN;
END_IF;

CheckInitialization := FRegistration.IsInitialized
    AND FOrder.IsInitialized
    AND FSlots.IsInitialized
    AND FFinalization.IsInitialized;
END_METHOD

{region 'Documentation'}
(*!
<summary>Configures one direct builder scenario and its named Assertions.</summary>
*)
{endregion}
METHOD PROTECTED Configure
FPreparationStateCount := 0;
FTestStateCount := 1;
FScenarioExecuted := FALSE;
FChecksEvaluated := FALSE;

FRegistrationMatches := FALSE;
FRegistration.Initialize(Parent := THIS^,
    AssertionName := 'Registration');
FOrderMatches := FALSE;
FOrder.Initialize(Parent := THIS^,
    AssertionName := 'Order');
FSlotsMatches := FALSE;
FSlots.Initialize(Parent := THIS^,
    AssertionName := 'Slots');
FFinalizationMatches := FALSE;
FFinalization.Initialize(Parent := THIS^,
    AssertionName := 'Finalization');
END_METHOD

{region 'Documentation'}
(*!
<summary>Completes Abort immediately; no asynchronous resource operation is started.</summary>
*)
{endregion}
METHOD PROTECTED ProcessAbort
VAR_INPUT
    Enable : BOOL; //! Phase permission supplied by the owning Test Case; FALSE does not authorize progression, while observation may continue.
END_VAR
IF Enable THEN
    CompleteAbort();
END_IF;
END_METHOD

{region 'Documentation'}
(*!
<summary>Evaluates recorded observations and consumes pending resets on disabled calls.</summary>
*)
{endregion}
METHOD PROTECTED ProcessAssertions
VAR_INPUT
    Enable : BOOL; //! Phase permission supplied by the owning Test Case; FALSE does not authorize progression, while observation may continue.
END_VAR
FRegistration(Enable := Enable,
    State := State,
    IN := FRegistrationMatches);

FOrder(Enable := Enable,
    State := State,
    IN := FOrderMatches);

FSlots(Enable := Enable,
    State := State,
    IN := FSlotsMatches);

FFinalization(Enable := Enable,
    State := State,
    IN := FFinalizationMatches);

IF Enable AND FRegistration.EvaluationActive
    AND FOrder.EvaluationActive
    AND FSlots.EvaluationActive
    AND FFinalization.EvaluationActive THEN
    FChecksEvaluated := TRUE;
END_IF;
END_METHOD

{region 'Documentation'}
(*!
<summary>No Preparation phase is needed for synchronous builder calls.</summary>
*)
{endregion}
METHOD PROTECTED ProcessPreparations
VAR_INPUT
    // SA0033: Required override signature; this scenario has no Preparation work.
    {attribute 'analysis' := '-33'}
    Enable : BOOL; //! Phase permission supplied by the owning Test Case; FALSE does not authorize progression, while observation may continue.
END_VAR
END_METHOD

{region 'Documentation'}
(*!
<summary>Clears recorded checks and Assertion results; each scenario initializes its own builder.</summary>
*)
{endregion}
METHOD PROTECTED ProcessReset
FScenarioExecuted := FALSE;
FChecksEvaluated := FALSE;
FRegistrationMatches := FALSE;
FRegistration.Reset();
FOrderMatches := FALSE;
FOrder.Reset();
FSlotsMatches := FALSE;
FSlots.Reset();
FFinalizationMatches := FALSE;
FFinalization.Reset();
CompleteReset();
END_METHOD

{region 'Documentation'}
(*!
<summary>Runs setup operations once, then completes after their observations have been evaluated.</summary>
*)
{endregion}
METHOD PROTECTED ProcessTests
VAR_INPUT
    Enable : BOOL; //! Phase permission supplied by the owning Test Case; FALSE does not authorize progression, while observation may continue.
END_VAR
IF NOT Enable THEN
    RETURN;
END_IF;

IF FChecksEvaluated THEN
    CompleteTests();
ELSIF NOT FScenarioExecuted THEN
    RunScenario();
    FScenarioExecuted := TRUE;
END_IF;
END_METHOD

{region 'Documentation'}
(*!
<summary>Checks stable insertion into two slots, including a temporary gap before Finalize.</summary>
*)
{endregion}
METHOD PRIVATE RunScenario
VAR
    ChildA : I_TestCase;
    ChildB : I_TestCase;
    ChildC : I_TestCase;
    ChildD : I_TestCase;
    AcceptedA : BOOL;
    AcceptedB : BOOL;
    AcceptedC : BOOL;
    AcceptedD : BOOL;
    Config : ST_TestCaseCollectionConfig;
END_VAR
ChildA := FChildA;
ChildB := FChildB;
ChildC := FChildC;
ChildD := FChildD;
FBuilder.Initialize(Mode := E_OrchestrationMode.ParallelSlots,
    TestCases := FCases);
AcceptedA := FBuilder.RegisterWithSlot(TestCase := ChildA,
    ExecutionSlot := 2);
AcceptedB := FBuilder.RegisterWithSlot(TestCase := ChildB,
    ExecutionSlot := 1);
AcceptedC := FBuilder.RegisterWithSlot(TestCase := ChildC,
    ExecutionSlot := 2);
AcceptedD := FBuilder.RegisterWithSlot(TestCase := ChildD,
    ExecutionSlot := 1);
FRegistrationMatches := AcceptedA AND AcceptedB AND AcceptedC AND AcceptedD;
FOrderMatches := (FCases[1] = ChildB) AND (FCases[2] = ChildD)
    AND (FCases[3] = ChildA) AND (FCases[4] = ChildC);
FSlotsMatches := (FChildA.ExecutionSlot = 2) AND (FChildB.ExecutionSlot = 1)
    AND (FChildC.ExecutionSlot = 2) AND (FChildD.ExecutionSlot = 1);

Config := FBuilder.Finalize();
FFinalizationMatches := Config.IsValid AND FBuilder.IsValid AND FBuilder.IsFinalized
    AND (Config.FirstIndex = 1) AND (Config.LastIndex = 4) AND (Config.Count = 4)
    AND (Config.Mode = E_OrchestrationMode.ParallelSlots);
END_METHOD

END_FUNCTION_BLOCK

// ---- SelfTests/TestCases/TestSuite_TestSuiteConfigurationBuilder/Test_SuiteBuilderCapacity.TcPOU
{region 'Documentation'}
(*!
<summary>Checks exact capacity and rejection before array or candidate-slot mutation.</summary>
<description>Child mocks are inert interface identities and slot storage only; no child initialization or FB call is performed.</description>
*)
{endregion}
FUNCTION_BLOCK Test_SuiteBuilderCapacity EXTENDS TestCaseBase
VAR
    FBuilder : TestSuiteConfigurationBuilder;
    FCases : ARRAY[1..2] OF I_TestCase;
    FChildA : TestCaseMock;
    FChildB : TestCaseMock;
    FChildC : TestCaseMock;
    FScenarioExecuted : BOOL;
    FChecksEvaluated : BOOL;
    FExactCapacity : AssertTrue;
    FExactCapacityMatches : BOOL;
    FOverflowRejected : AssertTrue;
    FOverflowRejectedMatches : BOOL;
    FCompositionPreserved : AssertTrue;
    FCompositionPreservedMatches : BOOL;
    FErrorLatched : AssertTrue;
    FErrorLatchedMatches : BOOL;
END_VAR
VAR CONSTANT
    CandidateSlotBeforeRejection : UINT := 9;
END_VAR

SUPER^();

{region 'Documentation'}
(*!
<summary>Contributes each owned Assertion once without executing it.</summary>
*)
{endregion}
METHOD PROTECTED AggregateResults
VAR_INPUT
    Aggregator : I_ResultAggregator; //! Borrowed result sink owned by the outer Test Case; add this test's checking Assertions without resetting or retaining the sink.
END_VAR
Aggregator.AddProvider(Provider := FExactCapacity);
Aggregator.AddProvider(Provider := FOverflowRejected);
Aggregator.AddProvider(Provider := FCompositionPreserved);
Aggregator.AddProvider(Provider := FErrorLatched);
END_METHOD

{region 'Documentation'}
(*!
<summary>Requires successful base and owned Assertion initialization.</summary>
*)
{endregion}
METHOD PROTECTED CheckInitialization : BOOL //! TRUE when the inherited initialization check and this concrete fixture check both accept the setup.
CheckInitialization := FALSE;
IF NOT SUPER^.CheckInitialization() THEN
    RETURN;
END_IF;

CheckInitialization := FExactCapacity.IsInitialized
    AND FOverflowRejected.IsInitialized
    AND FCompositionPreserved.IsInitialized
    AND FErrorLatched.IsInitialized;
END_METHOD

{region 'Documentation'}
(*!
<summary>Configures one direct builder scenario and its named Assertions.</summary>
*)
{endregion}
METHOD PROTECTED Configure
FPreparationStateCount := 0;
FTestStateCount := 1;
FScenarioExecuted := FALSE;
FChecksEvaluated := FALSE;

FExactCapacityMatches := FALSE;
FExactCapacity.Initialize(Parent := THIS^,
    AssertionName := 'ExactCapacity');
FOverflowRejectedMatches := FALSE;
FOverflowRejected.Initialize(Parent := THIS^,
    AssertionName := 'OverflowRejected');
FCompositionPreservedMatches := FALSE;
FCompositionPreserved.Initialize(Parent := THIS^,
    AssertionName := 'CompositionPreserved');
FErrorLatchedMatches := FALSE;
FErrorLatched.Initialize(Parent := THIS^,
    AssertionName := 'ErrorLatched');
END_METHOD

{region 'Documentation'}
(*!
<summary>Completes Abort immediately; no asynchronous resource operation is started.</summary>
*)
{endregion}
METHOD PROTECTED ProcessAbort
VAR_INPUT
    Enable : BOOL; //! Phase permission supplied by the owning Test Case; FALSE does not authorize progression, while observation may continue.
END_VAR
IF Enable THEN
    CompleteAbort();
END_IF;
END_METHOD

{region 'Documentation'}
(*!
<summary>Evaluates recorded observations and consumes pending resets on disabled calls.</summary>
*)
{endregion}
METHOD PROTECTED ProcessAssertions
VAR_INPUT
    Enable : BOOL; //! Phase permission supplied by the owning Test Case; FALSE does not authorize progression, while observation may continue.
END_VAR
FExactCapacity(Enable := Enable,
    State := State,
    IN := FExactCapacityMatches);

FOverflowRejected(Enable := Enable,
    State := State,
    IN := FOverflowRejectedMatches);

FCompositionPreserved(Enable := Enable,
    State := State,
    IN := FCompositionPreservedMatches);

FErrorLatched(Enable := Enable,
    State := State,
    IN := FErrorLatchedMatches);

IF Enable AND FExactCapacity.EvaluationActive
    AND FOverflowRejected.EvaluationActive
    AND FCompositionPreserved.EvaluationActive
    AND FErrorLatched.EvaluationActive THEN
    FChecksEvaluated := TRUE;
END_IF;
END_METHOD

{region 'Documentation'}
(*!
<summary>No Preparation phase is needed for synchronous builder calls.</summary>
*)
{endregion}
METHOD PROTECTED ProcessPreparations
VAR_INPUT
    // SA0033: Required override signature; this scenario has no Preparation work.
    {attribute 'analysis' := '-33'}
    Enable : BOOL; //! Phase permission supplied by the owning Test Case; FALSE does not authorize progression, while observation may continue.
END_VAR
END_METHOD

{region 'Documentation'}
(*!
<summary>Clears recorded checks and Assertion results; each scenario initializes its own builder.</summary>
*)
{endregion}
METHOD PROTECTED ProcessReset
FScenarioExecuted := FALSE;
FChecksEvaluated := FALSE;
FExactCapacityMatches := FALSE;
FExactCapacity.Reset();
FOverflowRejectedMatches := FALSE;
FOverflowRejected.Reset();
FCompositionPreservedMatches := FALSE;
FCompositionPreserved.Reset();
FErrorLatchedMatches := FALSE;
FErrorLatched.Reset();
CompleteReset();
END_METHOD

{region 'Documentation'}
(*!
<summary>Runs setup operations once, then completes after their observations have been evaluated.</summary>
*)
{endregion}
METHOD PROTECTED ProcessTests
VAR_INPUT
    Enable : BOOL; //! Phase permission supplied by the owning Test Case; FALSE does not authorize progression, while observation may continue.
END_VAR
IF NOT Enable THEN
    RETURN;
END_IF;

IF FChecksEvaluated THEN
    CompleteTests();
ELSIF NOT FScenarioExecuted THEN
    RunScenario();
    FScenarioExecuted := TRUE;
END_IF;
END_METHOD

{region 'Documentation'}
(*!
<summary>Checks exact capacity and rejection before array or candidate-slot mutation.</summary>
*)
{endregion}
METHOD PRIVATE RunScenario
VAR
    ChildA : I_TestCase;
    ChildB : I_TestCase;
    ChildC : I_TestCase;
    AcceptedA : BOOL;
    AcceptedB : BOOL;
    AcceptedC : BOOL;
    Config : ST_TestCaseCollectionConfig;
END_VAR
ChildA := FChildA;
ChildB := FChildB;
ChildC := FChildC;
FBuilder.Initialize(Mode := E_OrchestrationMode.Serial,
    TestCases := FCases);
AcceptedA := FBuilder.Register(TestCase := ChildA);
AcceptedB := FBuilder.Register(TestCase := ChildB);
Config := FBuilder.Finalize();
FExactCapacityMatches := AcceptedA AND AcceptedB AND Config.IsValid
    AND (Config.Count = 2) AND (FCases[1] = ChildA) AND (FCases[2] = ChildB);

FBuilder.Initialize(Mode := E_OrchestrationMode.Serial,
    TestCases := FCases);
AcceptedA := FBuilder.Register(TestCase := ChildA);
AcceptedB := FBuilder.Register(TestCase := ChildB);
FChildC.ExecutionSlot := CandidateSlotBeforeRejection;
AcceptedC := FBuilder.Register(TestCase := ChildC);
FOverflowRejectedMatches := AcceptedA AND AcceptedB AND NOT AcceptedC;
FCompositionPreservedMatches := (FBuilder.Count = 2)
    AND (FCases[1] = ChildA) AND (FCases[2] = ChildB)
    AND (FChildA.ExecutionSlot = 1) AND (FChildB.ExecutionSlot = 2)
    AND (FChildC.ExecutionSlot = CandidateSlotBeforeRejection);

Config := FBuilder.Finalize();
FErrorLatchedMatches := NOT Config.IsValid AND NOT FBuilder.IsValid
    AND FBuilder.IsFinalized AND (Config.Count = 2);
END_METHOD

END_FUNCTION_BLOCK

// ---- SelfTests/TestCases/TestSuite_TestSuiteConfigurationBuilder/Test_SuiteBuilderRegistrationErrors.TcPOU
{region 'Documentation'}
(*!
<summary>Checks typical setup mistakes without executing the registered child objects.</summary>
<description>Child mocks are inert interface identities and slot storage only; no child initialization or FB call is performed.</description>
*)
{endregion}
FUNCTION_BLOCK Test_SuiteBuilderRegistrationErrors EXTENDS TestCaseBase
VAR
    FBuilder : TestSuiteConfigurationBuilder;
    FCases : ARRAY[1..2] OF I_TestCase;
    FChildA : TestCaseMock;
    FChildB : TestCaseMock;
    FScenarioExecuted : BOOL;
    FChecksEvaluated : BOOL;
    FDuplicateRejected : AssertTrue;
    FDuplicateRejectedMatches : BOOL;
    FNullRejected : AssertTrue;
    FNullRejectedMatches : BOOL;
    FExplicitSlotRejected : AssertTrue;
    FExplicitSlotRejectedMatches : BOOL;
    FMissingSlotRejected : AssertTrue;
    FMissingSlotRejectedMatches : BOOL;
    FZeroSlotRejected : AssertTrue;
    FZeroSlotRejectedMatches : BOOL;
    FSlotGapRejected : AssertTrue;
    FSlotGapRejectedMatches : BOOL;
END_VAR
VAR CONSTANT
    CandidateSlotBeforeRejection : UINT := 9;
END_VAR

SUPER^();

{region 'Documentation'}
(*!
<summary>Contributes each owned Assertion once without executing it.</summary>
*)
{endregion}
METHOD PROTECTED AggregateResults
VAR_INPUT
    Aggregator : I_ResultAggregator; //! Borrowed result sink owned by the outer Test Case; add this test's checking Assertions without resetting or retaining the sink.
END_VAR
Aggregator.AddProvider(Provider := FDuplicateRejected);
Aggregator.AddProvider(Provider := FNullRejected);
Aggregator.AddProvider(Provider := FExplicitSlotRejected);
Aggregator.AddProvider(Provider := FMissingSlotRejected);
Aggregator.AddProvider(Provider := FZeroSlotRejected);
Aggregator.AddProvider(Provider := FSlotGapRejected);
END_METHOD

{region 'Documentation'}
(*!
<summary>Requires successful base and owned Assertion initialization.</summary>
*)
{endregion}
METHOD PROTECTED CheckInitialization : BOOL //! TRUE when the inherited initialization check and this concrete fixture check both accept the setup.
CheckInitialization := FALSE;
IF NOT SUPER^.CheckInitialization() THEN
    RETURN;
END_IF;

CheckInitialization := FDuplicateRejected.IsInitialized
    AND FNullRejected.IsInitialized
    AND FExplicitSlotRejected.IsInitialized
    AND FMissingSlotRejected.IsInitialized
    AND FZeroSlotRejected.IsInitialized
    AND FSlotGapRejected.IsInitialized;
END_METHOD

{region 'Documentation'}
(*!
<summary>Configures one direct builder scenario and its named Assertions.</summary>
*)
{endregion}
METHOD PROTECTED Configure
FPreparationStateCount := 0;
FTestStateCount := 1;
FScenarioExecuted := FALSE;
FChecksEvaluated := FALSE;

FDuplicateRejectedMatches := FALSE;
FDuplicateRejected.Initialize(Parent := THIS^,
    AssertionName := 'DuplicateRejected');
FNullRejectedMatches := FALSE;
FNullRejected.Initialize(Parent := THIS^,
    AssertionName := 'NullRejected');
FExplicitSlotRejectedMatches := FALSE;
FExplicitSlotRejected.Initialize(Parent := THIS^,
    AssertionName := 'ExplicitSlotRejected');
FMissingSlotRejectedMatches := FALSE;
FMissingSlotRejected.Initialize(Parent := THIS^,
    AssertionName := 'MissingSlotRejected');
FZeroSlotRejectedMatches := FALSE;
FZeroSlotRejected.Initialize(Parent := THIS^,
    AssertionName := 'ZeroSlotRejected');
FSlotGapRejectedMatches := FALSE;
FSlotGapRejected.Initialize(Parent := THIS^,
    AssertionName := 'SlotGapRejected');
END_METHOD

{region 'Documentation'}
(*!
<summary>Completes Abort immediately; no asynchronous resource operation is started.</summary>
*)
{endregion}
METHOD PROTECTED ProcessAbort
VAR_INPUT
    Enable : BOOL; //! Phase permission supplied by the owning Test Case; FALSE does not authorize progression, while observation may continue.
END_VAR
IF Enable THEN
    CompleteAbort();
END_IF;
END_METHOD

{region 'Documentation'}
(*!
<summary>Evaluates recorded observations and consumes pending resets on disabled calls.</summary>
*)
{endregion}
METHOD PROTECTED ProcessAssertions
VAR_INPUT
    Enable : BOOL; //! Phase permission supplied by the owning Test Case; FALSE does not authorize progression, while observation may continue.
END_VAR
FDuplicateRejected(Enable := Enable,
    State := State,
    IN := FDuplicateRejectedMatches);

FNullRejected(Enable := Enable,
    State := State,
    IN := FNullRejectedMatches);

FExplicitSlotRejected(Enable := Enable,
    State := State,
    IN := FExplicitSlotRejectedMatches);

FMissingSlotRejected(Enable := Enable,
    State := State,
    IN := FMissingSlotRejectedMatches);

FZeroSlotRejected(Enable := Enable,
    State := State,
    IN := FZeroSlotRejectedMatches);

FSlotGapRejected(Enable := Enable,
    State := State,
    IN := FSlotGapRejectedMatches);

IF Enable AND FDuplicateRejected.EvaluationActive
    AND FNullRejected.EvaluationActive
    AND FExplicitSlotRejected.EvaluationActive
    AND FMissingSlotRejected.EvaluationActive
    AND FZeroSlotRejected.EvaluationActive
    AND FSlotGapRejected.EvaluationActive THEN
    FChecksEvaluated := TRUE;
END_IF;
END_METHOD

{region 'Documentation'}
(*!
<summary>No Preparation phase is needed for synchronous builder calls.</summary>
*)
{endregion}
METHOD PROTECTED ProcessPreparations
VAR_INPUT
    // SA0033: Required override signature; this scenario has no Preparation work.
    {attribute 'analysis' := '-33'}
    Enable : BOOL; //! Phase permission supplied by the owning Test Case; FALSE does not authorize progression, while observation may continue.
END_VAR
END_METHOD

{region 'Documentation'}
(*!
<summary>Clears recorded checks and Assertion results; each scenario initializes its own builder.</summary>
*)
{endregion}
METHOD PROTECTED ProcessReset
FScenarioExecuted := FALSE;
FChecksEvaluated := FALSE;
FDuplicateRejectedMatches := FALSE;
FDuplicateRejected.Reset();
FNullRejectedMatches := FALSE;
FNullRejected.Reset();
FExplicitSlotRejectedMatches := FALSE;
FExplicitSlotRejected.Reset();
FMissingSlotRejectedMatches := FALSE;
FMissingSlotRejected.Reset();
FZeroSlotRejectedMatches := FALSE;
FZeroSlotRejected.Reset();
FSlotGapRejectedMatches := FALSE;
FSlotGapRejected.Reset();
CompleteReset();
END_METHOD

{region 'Documentation'}
(*!
<summary>Runs setup operations once, then completes after their observations have been evaluated.</summary>
*)
{endregion}
METHOD PROTECTED ProcessTests
VAR_INPUT
    Enable : BOOL; //! Phase permission supplied by the owning Test Case; FALSE does not authorize progression, while observation may continue.
END_VAR
IF NOT Enable THEN
    RETURN;
END_IF;

IF FChecksEvaluated THEN
    CompleteTests();
ELSIF NOT FScenarioExecuted THEN
    RunScenario();
    FScenarioExecuted := TRUE;
END_IF;
END_METHOD

{region 'Documentation'}
(*!
<summary>Checks typical setup mistakes without executing the registered child objects.</summary>
*)
{endregion}
METHOD PRIVATE RunScenario
VAR
    ChildA : I_TestCase;
    ChildB : I_TestCase;
    AcceptedA : BOOL;
    AcceptedB : BOOL;
    Config : ST_TestCaseCollectionConfig;
    AcceptedAfterError : BOOL;
END_VAR
ChildA := FChildA;
ChildB := FChildB;
FBuilder.Initialize(Mode := E_OrchestrationMode.Serial,
    TestCases := FCases);
AcceptedA := FBuilder.Register(TestCase := ChildA);
AcceptedB := FBuilder.Register(TestCase := ChildA);
AcceptedAfterError := FBuilder.Register(TestCase := ChildB);
Config := FBuilder.Finalize();
FDuplicateRejectedMatches := AcceptedA AND NOT AcceptedB AND NOT AcceptedAfterError
    AND NOT Config.IsValid AND (FBuilder.Count = 1)
    AND (FCases[1] = ChildA) AND (FCases[2] = 0) AND (FChildA.ExecutionSlot = 1);

FBuilder.Initialize(Mode := E_OrchestrationMode.Serial,
    TestCases := FCases);
AcceptedA := FBuilder.Register(TestCase := ChildA);
AcceptedB := FBuilder.Register(TestCase := 0);
Config := FBuilder.Finalize();
FNullRejectedMatches := AcceptedA AND NOT AcceptedB AND NOT Config.IsValid
    AND (FBuilder.Count = 1) AND (FCases[1] = ChildA) AND (FCases[2] = 0);

FBuilder.Initialize(Mode := E_OrchestrationMode.Serial,
    TestCases := FCases);
FChildA.ExecutionSlot := CandidateSlotBeforeRejection;
AcceptedA := FBuilder.RegisterWithSlot(TestCase := ChildA,
    ExecutionSlot := 1);
Config := FBuilder.Finalize();
FExplicitSlotRejectedMatches := NOT AcceptedA AND NOT Config.IsValid
    AND (FBuilder.Count = 0) AND (FCases[1] = 0)
    AND (FChildA.ExecutionSlot = CandidateSlotBeforeRejection);

FBuilder.Initialize(Mode := E_OrchestrationMode.ParallelSlots,
    TestCases := FCases);
AcceptedA := FBuilder.Register(TestCase := ChildA);
Config := FBuilder.Finalize();
FMissingSlotRejectedMatches := NOT AcceptedA AND NOT Config.IsValid
    AND (FBuilder.Count = 0) AND (FCases[1] = 0)
    AND (FChildA.ExecutionSlot = CandidateSlotBeforeRejection);

